(* IEC 61131-3 sources: plcassist-cli/packages/volt-lsp-iec/test-corpus/awa-palletizer/Device/Plc Logic/Application/Library Manager/L_TS2P_TechModulesSynchronizingCamming, 102 files *)

(* ---- L_TS2P_INTERNAL.gvl ---- *)
VAR_GLOBAL
	CDIENUMSTARTVALUE : DINT := 22000;
END_VAR

(* ---- L_TS2M_ITFFLYINGSAWSTATEFMDATA.itf ---- *)
INTERFACE L_TS2M_ITFFLYINGSAWSTATEFMDATA
END_INTERFACE

(* ---- L_TS2M_ITFFLYINGSAWSTATETMDATA.itf ---- *)
INTERFACE L_TS2M_ITFFLYINGSAWSTATETMDATA
END_INTERFACE

METHOD MOVETOPARKPOS : BOOL
VAR_INPUT
	XEXECUTEMOVETOPARKPOS : BOOL;
	LRPARKPOSITION : LREAL := 180;
	EPOSITIONINGDIRECTION : MC_DIRECTION := MC_DIRECTION.mcPositiveDirection;
	LRPOSITIONINGVEL : LREAL := 10;
	LRPOSITIONINGACC : LREAL := 100;
	LRPOSITIONINGDEC : LREAL := 100;
	LRJERK : LREAL := 0;
END_VAR
VAR_OUTPUT
	XBUSY : BOOL;
	XDONE : BOOL;
	XCOMMANDABORTED : BOOL;
END_VAR
VAR_IN_OUT
	AXIS : AXIS_REF;
END_VAR
END_METHOD

(* ---- L_TS2P_ICONNECTORFLEXCAM.itf ---- *)
INTERFACE L_TS2P_ICONNECTORFLEXCAM
END_INTERFACE

(* ---- L_TS2P_ICONNECTORFLYINGSAW.itf ---- *)
INTERFACE L_TS2P_ICONNECTORFLYINGSAW
END_INTERFACE

(* ---- L_TS2P_ICONNECTORSYNCANDCORRECTION.itf ---- *)
INTERFACE L_TS2P_ICONNECTORSYNCANDCORRECTION
END_INTERFACE

(* ---- L_TS2P_ICONNECTORSYNCPOS.itf ---- *)
INTERFACE L_TS2P_ICONNECTORSYNCPOS
END_INTERFACE

(* ---- L_TS2P_IFLEXCAM.itf ---- *)
INTERFACE L_TS2P_IFLEXCAM
END_INTERFACE

METHOD CAM
VAR_INPUT
	ITFTECHMODULE : L_TS2P_IFlexCam;
	XENABLE : BOOL;
	XSYNCCAM : BOOL;
	SCCAMTABLE : MC_CAM_REF;
	LRCYCMASTERPOS : LREAL;
	LRCYCMASTERVEL : LREAL;
	LRCYCMASTERACC : LREAL;
	LRSLAVEPOS : LREAL;
	LRSLAVEVEL : LREAL;
	LRSLAVEACC : LREAL;
	EOFFSETMODEMASTER : L_TS2P_OffsetMode := L_TS2P_OffsetMode.x_zero;
	ESCALINGMODEMASTER : L_TS2P_ScalingMode := L_TS2P_ScalingMode.x_zero;
	EOFFSETMODESLAVE : L_TS2P_OffsetMode := L_TS2P_OffsetMode.x_zero;
	ESCALINGMODESLAVE : L_TS2P_ScalingMode := L_TS2P_ScalingMode.x_zero;
	LRSETOFFSETMASTER : LREAL;
	LRSETOFFSETSLAVE : LREAL;
	LRSETSCALINGMASTER : LREAL;
	LRSETSCALINGSLAVE : LREAL;
	LRPROFGENMASTERVEL : LREAL;
	LRPROFGENMASTERACC : LREAL;
	LRPROFGENMASTERDEC : LREAL;
	LRPROFGENMASTERJERK : LREAL;
	LRPROFGENSLAVEVEL : LREAL;
	LRPROFGENSLAVEACC : LREAL;
	LRPROFGENSLAVEDEC : LREAL;
	LRPROFGENSLAVEJERK : LREAL;
	XPERIODIC : BOOL;
	XCAMCHANGEINSTANT : BOOL;
	XMASTERABSOLUTE : BOOL;
	XSLAVEABSOLUTE : BOOL;
END_VAR
VAR_OUTPUT
	XERROR : BOOL;
	EERRORID : L_IE1P.L_IE1P_Error;
	LRSETPOSOUT : LREAL;
	LRSETVELOUT : LREAL;
	LRSETACCOUT : LREAL;
	LRSETXPOSOUT : LREAL;
	LRSETXVELOUT : LREAL;
	LRSETXACCOUT : LREAL;
	LRSETYPOSOUT : LREAL;
	LRSETYVELOUT : LREAL;
	LRSETYACCOUT : LREAL;
	XENDOFPROFILE : BOOL;
	LRSETOFFSETMASTEROUT : LREAL;
	LRSETOFFSETSLAVEOUT : LREAL;
	LRCONVERTMASTERTOXPOS : LREAL;
	LRCAMPROFILERPOSOUT : LREAL;
	LRCONVERTYTOSLAVEPOS : LREAL;
	XDONE : BOOL;
	XBUSY : BOOL;
END_VAR
END_METHOD

METHOD CAMSEQUENCER
VAR_INPUT
	ITFTECHMODULE : L_TS2P_IFlexCam;
	XENABLE : BOOL;
	XCAMSEQUENCER : BOOL;
	XENDOFPROFILEIN : BOOL;
	CAMTABLE1 : MC_CAM_REF;
	CAMTABLE2 : MC_CAM_REF;
	CAMTABLE3 : MC_CAM_REF;
	CAMTABLE4 : MC_CAM_REF;
	XCAMCHANGEINSTANT : BOOL;
	XLOADCAMTABLE : BOOL;
	WSETCAMTABLE : WORD;
	EMODE : L_TS2P_CamSequenceMode := L_TS2P_CamSequenceMode.CyclicCam1;
END_VAR
VAR_OUTPUT
	XERROR : BOOL;
	EERRORID : L_IE1P_Error;
	CAMTABLEOUT : MC_CAM_REF;
	XCAMTABLEVALID : BOOL;
END_VAR
END_METHOD

METHOD CLUTCH
VAR_INPUT
	ITFTECHMODULE : L_TS2P_IFlexCam;
	XENABLE : BOOL;
	XCLUTCHCLOSE : BOOL;
	ECLUTCHINMODE : L_TS2P_ClutchInMode;
	ECLUTCHOUTMODE : L_TS2P_ClutchOutMode;
	EALLOWEDDIRECTION : L_TB2P_AllowedDirection;
	LRCLUTCHINDIST : LREAL;
	LRCLUTCHOUTDIST : LREAL;
	LRCLUTCHOUTPOSITION : LREAL;
	LRCYCLICMASTERPOS : LREAL;
	LRCYCLICMASTERVEL : LREAL;
	LRCYCLICMASTERACC : LREAL;
	LRCYCLICAXISPOS : LREAL;
	LRCYCLICAXISVEL : LREAL;
	LRCYCLICAXISACC : LREAL;
	ETRAVERSINGRANGE : L_MC1P_TraversingRange;
	LRCYCLELENGTH : LREAL;
END_VAR
VAR_OUTPUT
	XERROR : BOOL;
	EERRORID : L_IE1P.L_IE1P_Error;
	XBUSY : BOOL;
	XDONE : BOOL;
	XSYNCHRONISED : BOOL;
	XACCDECSYNC : BOOL;
	LRSETPOSOUT : LREAL;
	LRSETVELOUT : LREAL;
	LRSETACCOUT : LREAL;
END_VAR
END_METHOD

METHOD HALT : BOOL
VAR_INPUT
	ITFTECHMODULE : L_TS2P_IFlexCam;
	XEXECUTE : BOOL;
	LRDEC : LREAL := 100;
	LRJERK : LREAL := 0;
END_VAR
VAR_OUTPUT
	XBUSY : BOOL;
	XDONE : BOOL;
	XCOMMANDABORTED : BOOL;
END_VAR
VAR_IN_OUT
	AXIS : AXIS_REF;
END_VAR
END_METHOD

METHOD MOVETOPARKPOS : BOOL
VAR_INPUT
	ITFTECHMODULE : L_TS2P_IFlexCam;
	XEXECUTEMOVETOPARKPOS : BOOL;
	EMOVETOPARKPOSMODE : L_TS2P_CamStopMode;
	LRPARKPOSITION : LREAL := 180;
	EPOSITIONINGDIRECTION : L_TS2P_SyncDirection := L_TS2P_SyncDirection.PositiveDirection;
	LRPOSITIONINGVEL : LREAL := 10;
	LRPOSITIONINGACC : LREAL := 100;
	LRPOSITIONINGDEC : LREAL := 100;
	LRJERK : LREAL := 0;
END_VAR
VAR_OUTPUT
	XBUSY : BOOL;
	XDONE : BOOL;
	XCOMMANDABORTED : BOOL;
END_VAR
VAR_IN_OUT
	AXIS : AXIS_REF;
END_VAR
END_METHOD

METHOD POSITIONFOLLOWER
VAR_INPUT
	ITFTECHMODULE : L_TS2P_IFlexCam;
	XENABLE : BOOL;
	LRPOSITION : LREAL;
	LRVELOCITY : LREAL;
	LRACCELERATION : LREAL;
	ESETVALUEMODE : L_MC1P_SetValueMode;
END_VAR
VAR_OUTPUT
	XERROR : BOOL;
	EERRORID : L_IE1P.L_IE1P_Error;
	XBUSY : BOOL;
END_VAR
END_METHOD

METHOD SYNCIN
VAR_INPUT
	ITFTECHMODULE : L_TS2P_IFlexCam;
	XENABLE : BOOL;
	XSYNCIN : BOOL;
	XSYNCPOSRESTORE : BOOL;
	ESYNCMODE : L_TS2P_SyncInMode;
	ESYNCDIRECTION : L_TS2P_SyncDirection;
	LRSYNCVEL : LREAL;
	LRSYNCACC : LREAL;
	LRSYNCDEC : LREAL;
	LRSYNCJERK : LREAL;
	LRPARKPOSITION : LREAL;
	LRCYCLICMASTERPOS : LREAL;
	LRCYCLICMASTERVEL : LREAL;
	LRCYCLICMASTERACC : LREAL;
	LRCYCLICAXISPOS : LREAL;
	LRCYCLICAXISVEL : LREAL;
	LRCYCLICAXISACC : LREAL;
END_VAR
VAR_OUTPUT
	XERROR : BOOL;
	EERRORID : L_IE1P.L_IE1P_Error;
	XBUSY : BOOL;
	XDONE : BOOL;
	XSYNCHRONISED : BOOL;
	XACCDECSYNC : BOOL;
	LRSETPOSOUT : LREAL;
	LRSETVELOUT : LREAL;
	LRSETACCOUT : LREAL;
	LROFFSETSYNCPOS : LREAL;
END_VAR
VAR_IN_OUT
	AXIS : AXIS_REF;
END_VAR
END_METHOD

(* ---- L_TS2P_IFLYINGSAWPROCESSING.itf ---- *)
INTERFACE L_TS2P_IFLYINGSAWPROCESSING
END_INTERFACE

METHOD CLUTCH
VAR_INPUT
	ITFTECHMODULE : L_TS2P_IFlyingSawProcessing;
	XENABLE : BOOL;
	XSYNCVEL : BOOL := FALSE;
	XSYNCPOS : BOOL;
	XSYNCOUTINSTANT : BOOL;
	LRSYNCVEL : LREAL := 10;
	LRSYNCACC : LREAL := 100;
	LRSYNCDEC : LREAL := 100;
	LRSYNCJERK : LREAL := 10000;
	LRCYCMASTERPOS : LREAL;
	LRCYCMASTERVEL : LREAL;
	LRCYCMASTERACC : LREAL;
	LRSETSLAVEPOS : LREAL;
	LRSETSLAVEVEL : LREAL;
	LRSETSLAVEACC : LREAL;
END_VAR
VAR_OUTPUT
	EERRORID : L_IE1P_Error;
	XERROR : BOOL;
	XBUSY : BOOL;
	XDONE : BOOL;
	XACCDECSYNC : BOOL;
	XVELSYNCHRONISED : BOOL;
	XPOSSYNCHRONISED : BOOL;
	LRSETSLAVEPOSOUT : LREAL;
	LRSETSLAVEVELOUT : LREAL;
	LRSETSLAVEACCOUT : LREAL;
	XPROFILERESETTIMEVALID : BOOL;
	LRPROFILERESETTIME : LREAL;
END_VAR
END_METHOD

METHOD EXECUTEGAP
VAR_INPUT
	ITFTECHMODULE : L_TS2P_IFlyingSawProcessing;
	XENABLE : BOOL;
	LRSYNCVEL : LREAL := 10;
	LRSYNCACC : LREAL := 100;
	LRSYNCDEC : LREAL := 100;
	LRSYNCJERK : LREAL := 10000;
	XEXECUTEGAP : BOOL;
	XAUXEXECUTEGAP : BOOL := FALSE;
	LRCYCMASTERPOS : LREAL;
	LRCYCMASTERVEL : LREAL;
	LRCYCMASTERACC : LREAL;
	LRSETSLAVEPOS : LREAL;
	LRSETSLAVEVEL : LREAL;
	LRSETSLAVEACC : LREAL;
END_VAR
VAR_OUTPUT
	EERRORID : L_IE1P_Error;
	XERROR : BOOL;
	XBUSY : BOOL;
	XDONE : BOOL;
	XACCDECSYNC : BOOL;
	XVELSYNCHRONISED : BOOL;
	XPOSSYNCHRONISED : BOOL;
	LRSETSLAVEPOSOUT : LREAL;
	LRSETSLAVEVELOUT : LREAL;
	LRSETSLAVEACCOUT : LREAL;
	XPROFILERESETTIMEVALID : BOOL;
	LRPROFILERESETTIME : LREAL;
END_VAR
END_METHOD

METHOD MARKSTACK_GETMARK
VAR_INPUT
	ITFTECHMODULE : L_TS2P_IFlyingSawProcessing;
	XENABLE : BOOL;
	XGETMARK : BOOL;
	XRESETGETMARK : BOOL;
	XRESETMARKSTACK : BOOL;
	LRCYCSETPOS : LREAL;
	LRCYCSETVEL : LREAL;
END_VAR
VAR_OUTPUT
	XMARKSTACKFULL : BOOL;
	XMARKSTACKEMPTY : BOOL;
	WMARKSINSTACK : WORD;
	XMARKVALID : BOOL;
	LRMARKPOSOUT : LREAL;
END_VAR
END_METHOD

METHOD MARKSTACK_SETMARK
VAR_INPUT
	ITFTECHMODULE : L_TS2P_IFlyingSawProcessing;
	XENABLE : BOOL;
	XSETMARK : BOOL;
	LRMARKPOS : LREAL;
	XRESETMARKSTACK : BOOL;
	LRCYCSETPOS : LREAL;
	LRCYCSETVEL : LREAL;
END_VAR
VAR_OUTPUT
	XMARKSTACKFULL : BOOL;
	XMARKSTACKEMPTY : BOOL;
	WMARKSINSTACK : WORD;
	XNEWMARKRECEIVED : BOOL;
END_VAR
END_METHOD

METHOD POSITIONING
VAR_INPUT
	ITFTECHMODULE : L_TS2P_IFlyingSawProcessing;
	XENABLE : BOOL;
	XMOVETOTARGETPOS : BOOL;
	LRTARGETPOS : LREAL;
	LRPOSITIONINGVEL : LREAL;
	LRPOSITIONINGACC : LREAL;
	LRPOSITIONINGDEC : LREAL;
	LRPOSITIONINGJERK : LREAL;
	LRSETSLAVEPOS : LREAL;
	LRSETSLAVEVEL : LREAL;
	LRSETSLAVEACC : LREAL;
	LRCORRECTTIMEBASE : LREAL := 0;
	LROVERRIDE : LREAL := 1.0;
END_VAR
VAR_OUTPUT
	EERRORID : L_IE1P_Error;
	XERROR : BOOL;
	XBUSY : BOOL;
	XDONE : BOOL;
	XPOSITIONING : BOOL;
	XINPOSITION : BOOL;
	LRSETSLAVEPOSOUT : LREAL;
	LRSETSLAVEVELOUT : LREAL;
	LRSETSLAVEACCOUT : LREAL;
	XPROFILERESETTIMEVALID : BOOL;
	LRPROFILERESETTIME : LREAL;
END_VAR
END_METHOD

(* ---- L_TS2P_ISIGNALFLOW.itf ---- *)
INTERFACE L_TS2P_ISIGNALFLOW
END_INTERFACE

METHOD GET_PSF : POINTER TO L_TS2P_scSF_TM_SyncPosBase
END_METHOD

(* ---- L_TS2P_ISIGNALFLOWFLEXCAM.itf ---- *)
INTERFACE L_TS2P_ISIGNALFLOWFLEXCAM
END_INTERFACE

METHOD GET_PSF : POINTER TO L_TS2P_scSF_TM_SyncPosBase
END_METHOD

(* ---- L_TS2P_ISIGNALFLOWSC.itf ---- *)
INTERFACE L_TS2P_ISIGNALFLOWSC
END_INTERFACE

METHOD GET_PSF : POINTER TO L_TS2P_scSF_TM_SyncAndCorrectionState
END_METHOD

(* ---- L_TS2P_ISTRUCTPROVIDERFLEXCAMHIGH.itf ---- *)
INTERFACE L_TS2P_ISTRUCTPROVIDERFLEXCAMHIGH
END_INTERFACE

METHOD GET_PDATA : POINTER TO L_TS2P_scData_TM_FlexCam
END_METHOD

METHOD GET_PDATASP : POINTER TO L_TS2P_scData_TM_FlexCam
END_METHOD

(* ---- L_TS2P_ISTRUCTPROVIDERFLYINGSAW.itf ---- *)
INTERFACE L_TS2P_ISTRUCTPROVIDERFLYINGSAW
END_INTERFACE

METHOD GET_PDATA : POINTER TO L_TS2M_scData_FlyingSawState
END_METHOD

METHOD GET_PFMDATA : POINTER TO L_TS2M_scData_FM_FlyingSaw
END_METHOD

(* ---- L_TS2P_ISTRUCTPROVIDERSYNCANDCORRECTION.itf ---- *)
INTERFACE L_TS2P_ISTRUCTPROVIDERSYNCANDCORRECTION
END_INTERFACE

METHOD GET_PDATA : POINTER TO L_TS2P_scData_TM_SyncAndCorrectionState
END_METHOD

METHOD GET_PDATASP : POINTER TO L_TS2P_scData_TM_SyncPosBase
END_METHOD

(* ---- L_TS2P_ISTRUCTPROVIDERSYNCPOS.itf ---- *)
INTERFACE L_TS2P_ISTRUCTPROVIDERSYNCPOS
END_INTERFACE

METHOD GET_PDATA : POINTER TO L_TS2P_scData_TM_SyncPosBase
END_METHOD

(* ---- L_TS2P_ISYNCANDCORRECTIONSTATE.itf ---- *)
INTERFACE L_TS2P_ISYNCANDCORRECTIONSTATE
END_INTERFACE

(* ---- L_TS2P_ISYNCPOSBASE.itf ---- *)
INTERFACE L_TS2P_ISYNCPOSBASE
END_INTERFACE

METHOD ADDOFFSET
VAR_INPUT
	ITFTECHMODULE : L_TS2P_ISyncPosBase;
	LRSETPOS : LREAL;
	LRSETVEL : LREAL;
	LRSETOFFSET : LREAL;
	LRSETOFFSETVEL : LREAL;
	ETRAVERSINGRANGE : L_MC1P.L_MC1P_TraversingRange;
	LRCYCLELENGTH : LREAL;
END_VAR
VAR_OUTPUT
	XERROR : BOOL;
	EERRORID : L_IE1P.L_IE1P_Error;
	LRSETPOSOUT : LREAL;
	LRSETVELOUT : LREAL;
END_VAR
END_METHOD

METHOD CLUTCH
VAR_INPUT
	ITFTECHMODULE : L_TS2P_ISyncPosBase;
	XENABLE : BOOL;
	XSYNCIN : BOOL;
	LRSETBASEVELOCITY : LREAL;
	ESYNCMODE : L_TB2P_SyncMode;
	EALLOWEDDIRECTION : L_TB2P_AllowedDirection;
	LRSYNCVEL : LREAL;
	LRSYNCACC : LREAL;
	LRSYNCDEC : LREAL;
	LRSYNCJERK : LREAL;
	LRSYNCINDIST : LREAL;
	LRSYNCOUTDIST : LREAL;
	LRSYNCOUTPOS : LREAL;
	XLOADCLUTCHOFFSET : BOOL;
	LRLOADCLUTCHOFFSET : LREAL;
	LRCYCLICMASTERPOS : LREAL;
	LRCYCLICMASTERVEL : LREAL;
	ETRAVERSINGRANGEMASTER : L_MC1P_TraversingRange;
	LRCYCLELENGTHMASTER : LREAL;
	LRCYCLICAXISPOS : LREAL;
	LRCYCLICAXISVEL : LREAL;
	LRCYCLICAXISACC : LREAL;
	ETRAVERSINGRANGEAXIS : L_MC1P_TraversingRange;
	LRCYCLELENGTHAXIS : LREAL;
END_VAR
VAR_OUTPUT
	XERROR : BOOL;
	EERRORID : L_IE1P.L_IE1P_Error;
	XBUSY : BOOL;
	XDONE : BOOL;
	XSYNCHRONISED : BOOL;
	XACCDECSYNC : BOOL;
	XINBASEVELOCITY : BOOL;
	LRSETPOSOUT : LREAL;
	LRSETVELOUT : LREAL;
	LRSETACCOUT : LREAL;
	LRCLUTCHOFFSETOUT : LREAL;
END_VAR
END_METHOD

METHOD GEARBOX
VAR_INPUT
	ITFTECHMODULE : L_TS2P_ISyncPosBase;
	XENABLE : BOOL;
	LRSETPOSX : LREAL;
	LRSETVELX : LREAL;
	DWNUMERATOR : DWORD;
	DWDENOMINATOR : DWORD;
	LRCYCLELENGTHX : LREAL;
	LRCYCLELENGTHY : LREAL;
	ETRAVERSINGRANGEX : L_MC1P.L_MC1P_TraversingRange;
	ETRAVERSINGRANGEY : L_MC1P.L_MC1P_TraversingRange;
	XLOADGEARBOXPOS : BOOL;
	LRLOADGEARBOXPOS : LREAL;
END_VAR
VAR_OUTPUT
	XERROR : BOOL;
	EERRORID : L_IE1P.L_IE1P_Error;
	LRSETPOSOUT : LREAL;
	LRSETVELOUT : LREAL;
END_VAR
END_METHOD

METHOD OFFSETANDTRIM
VAR_INPUT
	ITFTECHMODULE : L_TS2P_ISyncPosBase;
	XENABLE : BOOL;
	LRSETOFFSET : LREAL;
	XTRIMPOS : BOOL;
	XTRIMNEG : BOOL;
	LRSETTRIMDISTANCE : LREAL;
	ETRIMMODE : L_TS2P_TrimMode;
	XLOADOFFSET : BOOL;
	XRESETTRIMOFFSET : BOOL;
	LRSETVEL : LREAL;
	LRSETACC : LREAL;
	LRSETDEC : LREAL;
	LRSETJERK : LREAL;
	WACTDIRECTION : WORD;
	EALLOWEDDIRECTION : L_TB2P.L_TB2P_AllowedDirection;
	LRCYCMASTERPOS : LREAL;
	LRCYCMASTERVEL : LREAL;
	LRCYCMASTERACC : LREAL;
END_VAR
VAR_OUTPUT
	XERROR : BOOL;
	EERRORID : L_IE1P.L_IE1P_Error;
	XBUSY : BOOL;
	XDONE : BOOL;
	LRSETOFFSETOUTTOTAL : LREAL;
	LRSETOFFSETOUTTOTALVEL : LREAL;
	LRSETOFFSETOUT : LREAL;
	LRSETOFFSETOUTTRIM : LREAL;
END_VAR
END_METHOD

(* ---- GETBOOLEANPROPERTY.fun ---- *)
FUNCTION GETBOOLEANPROPERTY : BOOL
VAR_INPUT
	STKEY : WSTRING;
END_VAR
END_FUNCTION

(* ---- GETCOMPANY.fun ---- *)
FUNCTION GETCOMPANY : WSTRING
END_FUNCTION

(* ---- GETNUMBERPROPERTY.fun ---- *)
FUNCTION GETNUMBERPROPERTY : DINT
VAR_INPUT
	STKEY : WSTRING;
END_VAR
END_FUNCTION

(* ---- GETTEXTPROPERTY.fun ---- *)
FUNCTION GETTEXTPROPERTY : WSTRING
VAR_INPUT
	STKEY : WSTRING;
END_VAR
END_FUNCTION

(* ---- GETTEXTPROPERTY2.fun ---- *)
FUNCTION GETTEXTPROPERTY2 : POINTER TO WSTRING
VAR_INPUT
	STKEY : WSTRING;
END_VAR
END_FUNCTION

(* ---- GETTITLE.fun ---- *)
FUNCTION GETTITLE : WSTRING
END_FUNCTION

(* ---- GETVERSION.fun ---- *)
FUNCTION GETVERSION : VERSION
END_FUNCTION

(* ---- GETVERSIONPROPERTY.fun ---- *)
FUNCTION GETVERSIONPROPERTY : VERSION
VAR_INPUT
	STKEY : WSTRING;
END_VAR
END_FUNCTION

(* ---- L_MB1P_CONVERTPOSTOMODULOPOS.fun ---- *)
FUNCTION L_MB1P_CONVERTPOSTOMODULOPOS : LREAL
VAR_INPUT
	LRPOS : LREAL;
	LRPERIOD : LREAL;
END_VAR
VAR_OUTPUT
	DIREVCOUNTER : DINT;
END_VAR
END_FUNCTION

(* ---- L_MB1P_CONVERTPOSTOMODULOPOSEXTENDED.fun ---- *)
FUNCTION L_MB1P_CONVERTPOSTOMODULOPOSEXTENDED : LREAL
VAR_INPUT
	LRPOS : LREAL;
	LRPERIOD : LREAL;
END_VAR
VAR_OUTPUT
	DIREVCOUNTER : DINT;
END_VAR
END_FUNCTION

(* ---- L_MB1P_CONVERTPOSTOMODULOPOSFMOD.fun ---- *)
FUNCTION L_MB1P_CONVERTPOSTOMODULOPOSFMOD : LREAL
VAR_INPUT
	LRPOS : LREAL;
	LRPERIOD : LREAL;
END_VAR
END_FUNCTION

(* ---- L_MB1P_HLPCALCKOEFPOLY5THORD.fun ---- *)
FUNCTION L_MB1P_HLPCALCKOEFPOLY5THORD : ARRAY [0..5] OF LREAL
VAR_INPUT
	LRYPOSSTART : LREAL;
	LRYVELSTART : LREAL;
	LRYACCSTART : LREAL;
	LRYPOSEND : LREAL;
	LRYVELEND : LREAL;
	LRYACCEND : LREAL;
END_VAR
VAR_OUTPUT
	ALRKOEF : ARRAY [0..5] OF LREAL;
END_VAR
END_FUNCTION

(* ---- L_MB1P_HLPCALCYOFPOLY5THORDBASE.fun ---- *)
FUNCTION L_MB1P_HLPCALCYOFPOLY5THORDBASE : LREAL
VAR_OUTPUT
	LRYPOSSCALED : LREAL;
END_VAR
VAR_IN_OUT
	LRXPOSSCALED : LREAL;
	ALRKOEF : ARRAY [0..5] OF LREAL;
END_VAR
END_FUNCTION

(* ---- L_MB1P_HLPCALCYOFPOLY5THORDSTATE.fun ---- *)
FUNCTION L_MB1P_HLPCALCYOFPOLY5THORDSTATE : LREAL
VAR_INPUT
	LRXPOSSTART : LREAL;
	LRXPOSEND : LREAL := 1;
	LRSETXPOS : LREAL;
	ALRKOEF : ARRAY [0..5] OF LREAL;
END_VAR
VAR_OUTPUT
	LRYPOSSCALED : LREAL;
END_VAR
END_FUNCTION

(* ---- L_MB1P_HLPDELTAVELTIMEEXTENDED.fun ---- *)
FUNCTION L_MB1P_HLPDELTAVELTIMEEXTENDED : BOOL
VAR_INPUT
	LRVELSTART : LREAL;
	LRACCSTART : LREAL;
	LRMAXACC : LREAL;
	LRMAXJERK : LREAL;
END_VAR
VAR_OUTPUT
	LRTIME : LREAL;
	LRDIST : LREAL;
END_VAR
END_FUNCTION

(* ---- L_MB1P_HLPDELTAVELTIMESTATE.fun ---- *)
FUNCTION L_MB1P_HLPDELTAVELTIMESTATE : BOOL
VAR_INPUT
	LRVELSTART : LREAL;
	LRACCSTART : LREAL;
	LRVELTARGET : LREAL;
	LRACCTARGET : LREAL;
	LRMAXACC : LREAL;
	LRMAXDEC : LREAL;
	LRMAXJERK : LREAL;
END_VAR
VAR_OUTPUT
	LRTIME : LREAL;
	LRDIST : LREAL;
END_VAR
END_FUNCTION

(* ---- L_MB1P_HLPDELTAVELTIMETOCONTANTVEL.fun ---- *)
FUNCTION L_MB1P_HLPDELTAVELTIMETOCONTANTVEL : BOOL
VAR_INPUT
	LRACCSTART : LREAL;
	LRMAXJERK : LREAL;
	WMODE : WORD;
END_VAR
VAR_OUTPUT
	LRVEL : LREAL;
	LRTIME : LREAL;
	LRDIST : LREAL;
END_VAR
END_FUNCTION

(* ---- L_MB1P_HLPRESTTIMEFORDISTANCE.fun ---- *)
FUNCTION L_MB1P_HLPRESTTIMEFORDISTANCE : BOOL
VAR_OUTPUT
	LRTIME : LREAL;
END_VAR
VAR_IN_OUT
	LRVELSTART : LREAL;
	LRACCSTART : LREAL;
	LRDIST : LREAL;
END_VAR
END_FUNCTION

(* ---- L_MB1P_MODULOCYCLE.fun ---- *)
FUNCTION L_MB1P_MODULOCYCLE : LREAL
VAR_INPUT
	LRPOSIN : LREAL;
	LRPOSITIONPERIOD : LREAL;
END_VAR
END_FUNCTION

(* ---- L_TS2P_CALCSYNCTIME.fun ---- *)
FUNCTION L_TS2P_CALCSYNCTIME : BOOL
VAR_INPUT
	LRACTMATERIALVEL : LREAL;
	LRACCMAX : LREAL;
	LRJERKSTART : LREAL;
	LRJERKEND : LREAL;
END_VAR
VAR_OUTPUT
	LRACCTIME : LREAL;
	LRACCDIST : LREAL;
END_VAR
END_FUNCTION

(* ---- L_TS2P_CHECK_CAMREFCHANGED.fun ---- *)
FUNCTION L_TS2P_CHECK_CAMREFCHANGED : BOOL
VAR_INPUT
	CAMREFNEW : MC_CAM_REF;
	CAMREFOLD : MC_CAM_REF;
END_VAR
END_FUNCTION

(* ---- L_TS2P_CHECK_CAMREFVALID.fun ---- *)
FUNCTION L_TS2P_CHECK_CAMREFVALID : BOOL
VAR_INPUT
	CAMREF : MC_CAM_REF;
END_VAR
END_FUNCTION

(* ---- _L_MB1P_AXISCONTROLBYPOS.fb ---- *)
FUNCTION_BLOCK _L_MB1P_AXISCONTROLBYPOS
VAR_INPUT
	XENABLE : BOOL;
	LRSETPOSITION : LREAL;
	LRSETVELOCITY : LREAL;
	LRSETACCELERATION : LREAL;
	ESETVALUEMODE : L_MC1P_SetValueMode := L_MC1P_SetValueMode.Pos;
END_VAR
VAR_OUTPUT
	XBUSY : BOOL;
	XCOMMANDABORTED : BOOL;
	XERROR : BOOL;
	EERRORID : L_IE1P_Error;
	LRSETPOSOUT : LREAL;
END_VAR
VAR_IN_OUT
	AXIS : AXIS_REF;
END_VAR
VAR
	LRSETPOSITION_INT : LREAL;
	XENABLE_OLD : BOOL;
	XBUSY_OLD : BOOL;
	ESTATE : L_MB1P_States;
	MC_HALT1 : MC_HALT;
	FB_FOLLOWSETVALUES : L_MC1P_FollowSetValues;
END_VAR
END_FUNCTION_BLOCK

METHOD CALL_ERRORHANDLER
END_METHOD

METHOD CALL_FBMETHODS
END_METHOD

METHOD CALL_FB_FOLLOWSETVALUES
END_METHOD

METHOD CALL_MC_HALT
END_METHOD

METHOD CALL_MC_HALT_INPUT
END_METHOD

METHOD CALL_OUTPUT
END_METHOD

METHOD CALL_RESETCOMMANDS
END_METHOD

METHOD CALL_RESETOUTPUT
END_METHOD

METHOD CALL_STATEMACHINE
END_METHOD

METHOD CALL_S000_CYCLIC
END_METHOD

METHOD CALL_S001_INIT
END_METHOD

METHOD CALL_S002_READY
END_METHOD

METHOD CALL_S999_ERROR
END_METHOD

(* ---- _L_MB1P_AXISCONTROLBYVEL.fb ---- *)
FUNCTION_BLOCK _L_MB1P_AXISCONTROLBYVEL
VAR_INPUT
	XENABLE : BOOL;
	LRSETVELOCITY : LREAL;
END_VAR
VAR_OUTPUT
	XBUSY : BOOL;
	XCOMMANDABORTED : BOOL;
	XERROR : BOOL;
	EERRORID : L_IE1P_Error;
	LRSETVELOUT : LREAL;
END_VAR
VAR_IN_OUT
	AXIS : AXIS_REF;
END_VAR
VAR
	LRSETVELOCITY_INT : LREAL;
	XENABLE_OLD : BOOL;
	XBUSY_OLD : BOOL;
	ESTATE : L_MB1P_States;
	MC_HALT1 : MC_HALT;
	FB_FOLLOWSETVALUES : L_MC1P_FollowSetValues;
END_VAR
END_FUNCTION_BLOCK

METHOD CALL_ERRORHANDLER
END_METHOD

METHOD CALL_FBMETHODS
END_METHOD

METHOD CALL_FB_FOLLOWSETVALUES
END_METHOD

METHOD CALL_MC_HALT
END_METHOD

METHOD CALL_MC_HALT_INPUT
END_METHOD

METHOD CALL_OUTPUT
END_METHOD

METHOD CALL_RESETCOMMANDS
END_METHOD

METHOD CALL_RESETOUTPUT
END_METHOD

METHOD CALL_STATEMACHINE
END_METHOD

METHOD CALL_S000_CYCLIC
END_METHOD

METHOD CALL_S001_INIT
END_METHOD

METHOD CALL_S002_READY
END_METHOD

METHOD CALL_S999_ERROR
END_METHOD

(* ---- GLOBALTEXTLIST.fb ---- *)
FUNCTION_BLOCK GLOBALTEXTLIST
VAR
	M_TEXTLISTFILE : STRING(255);
	_STNAMESPACE : STRING;
END_VAR
END_FUNCTION_BLOCK

(* ---- L_MB1P_CHECKMODULOOVERRUN.fb ---- *)
FUNCTION_BLOCK L_MB1P_CHECKMODULOOVERRUN
VAR_INPUT
	LRSETPOS : LREAL;
	LRSETVEL : LREAL;
	LRPERIOD : LREAL;
END_VAR
VAR_OUTPUT
	XOVERRUNPOS : BOOL;
	XOVERRUNNEG : BOOL;
END_VAR
VAR
	ALRMEM : ARRAY [1..7] OF LREAL;
END_VAR
END_FUNCTION_BLOCK

METHOD CALL_CHECKMODULOOVERRUN
VAR_IN_OUT
	LRSETPOS : LREAL;
	LRSETVEL : LREAL;
	LRPERIOD : LREAL;
	XOVERRUNPOS : BOOL;
	XOVERRUNNEG : BOOL;
	ALRMEM : ARRAY [1..7] OF LREAL;
END_VAR
END_METHOD

(* ---- L_MB1P_CHECKUNLIMITEDOVERRUN.fb ---- *)
FUNCTION_BLOCK L_MB1P_CHECKUNLIMITEDOVERRUN
VAR_INPUT
	LRSETPOS : LREAL;
	LRSETVEL : LREAL;
	LRPERIOD : LREAL;
END_VAR
VAR_OUTPUT
	XOVERRUNPOS : BOOL;
	XOVERRUNNEG : BOOL;
END_VAR
VAR
	ALRMEM : ARRAY [1..7] OF LREAL;
END_VAR
END_FUNCTION_BLOCK

METHOD CALL_CHECKUNLIMITEDOVERRUN
VAR_IN_OUT
	LRSETPOS : LREAL;
	LRSETVEL : LREAL;
	LRPERIOD : LREAL;
	XOVERRUNPOS : BOOL;
	XOVERRUNNEG : BOOL;
	ALRMEM : ARRAY [1..7] OF LREAL;
END_VAR
END_METHOD

(* ---- L_MB1P_CLUTCHEXTENDEDBASE.fb ---- *)
FUNCTION_BLOCK L_MB1P_CLUTCHEXTENDEDBASE EXTENDS L_MC2P_ClutchBasic
VAR_INPUT
	XENABLE : BOOL;
	XCLUTCHCLOSE : BOOL;
	XCLUTCHOPENINSTANT : BOOL;
	ECLUTCHMODE : L_MB1P_ClutchMode := L_MB1P_ClutchMode.ramp_pos;
	ECLUTCHDIRECTION : L_MC2P_ClutchDirection := L_MC2P_ClutchDirection.mcCurrentDirection;
	EDIRECTION : L_MC1P_Direction := 0;
	LRCYCMASTERPOS : LREAL;
	LRCYCMASTERVEL : LREAL;
	LRCYCMASTERACC : LREAL;
	LRCYCSLAVEPOS : LREAL;
	LRCYCSLAVEVEL : LREAL;
	LRCYCSLAVEACC : LREAL;
	LROPENINSTANTDEC : LREAL;
	LRMASTERCLOSEPOS : LREAL;
	LRMASTERCLOSEDIST : LREAL := 100;
	LRSLAVECLOSEDIST : LREAL := 100;
	LRMASTEROPENDIST : LREAL := 100;
	LRSLAVEOPENDIST : LREAL := 100;
	LRSLAVEOPENPOS : LREAL;
	LRCLOSETIME : LREAL := 5;
	LROPENTIME : LREAL := 5;
	LRCLUTCHVEL : LREAL := 100;
	LRCLUTCHACC : LREAL := 1000.0;
	LRCLUTCHDEC : LREAL := 1000.0;
	LRCLUTCHJERK : LREAL := 1000000.0;
	LRVELTOLERANCE : LREAL := 1;
	LRAXESCYCLELENGTH : LREAL := 360;
	EMASTERTRAVERSINGRANGE : L_MC1P_TraversingRange;
	LRCYCLETIME : LREAL := 0.001;
END_VAR
VAR_OUTPUT
	XERROR : BOOL;
	EERRORID : L_IE1P_Error;
	XBUSY : BOOL;
	XDONE : BOOL;
	XSYNCHRONISED : BOOL;
	XCLUTCHACTIVE : BOOL;
	LRSETSLAVEPOSOUT : LREAL;
	LRSETSLAVEVELOUT : LREAL;
	LRSETSLAVEACCOUT : LREAL;
	LRSETSLAVEOFFSETOUT : LREAL;
	LRX0 : LREAL;
	LRX1 : LREAL;
	LRY0 : LREAL;
	LRY1 : LREAL;
	LRX0N : LREAL;
	LRX1N : LREAL;
	LRY0N : LREAL;
	LRY1N : LREAL;
	LRX0P : LREAL;
	LRX1P : LREAL;
	LRY0P : LREAL;
	LRY1P : LREAL;
END_VAR
VAR
	EAXESTRAVERSINGRANGE_INT : L_MC1P_TraversingRange;
	ECLUTCHMODE_INT : L_MB1P_ClutchMode;
	ECLUTCHDIRECTION_INT : L_MB1P_ClutchDirection;
	LRSETSLAVEOFFSET_CLUTCHREL : LREAL;
	LRSETSLAVEOFFSET_INT : LREAL;
	LRSETMASTEROFFSET_OVERRUN : LREAL;
	LRCYCLETIME_INT : LREAL;
	XCLUTCHOPENINSTANT_ACTIVE : BOOL;
	LROPENINSTANTDEC_INT : LREAL;
	XCLUTCHBASICENABLE : BOOL;
	LRTEMP : LREAL;
	LRDELTASETENDPOS : LREAL;
	LRDELTASETENDPOS_OLD : LREAL;
	LRDELTASETENDPOS_OLD2 : LREAL;
	XCLUTCHMASTERVELPOSITIVE : BOOL;
	XMASTERREVERSING : BOOL;
	XCLUTCHBASIC_EXECUTE_OLD : BOOL;
	XCLUTCHCLOSE_OLD : BOOL;
	XCLUTCHOPENINSTANT_OLD : BOOL;
	XBUSY_OLD : BOOL;
	XENABLE_OLD : BOOL;
	LRCYCMASTERPOS_OLD : LREAL;
	LRMASTERVELADD : LREAL;
	LRMASTERVELADDSYNC : LREAL;
	LRSLAVESTARTPOS : LREAL;
	LRMASTERCLOSEPOS_INT : LREAL;
	LRMASTERCLOSEDIST_INT : LREAL;
	LRSLAVECLOSEDIST_INT : LREAL;
	LRSLAVEOPENDIST_INT : LREAL;
	LRSLAVEOPENPOS_INT : LREAL;
	XSYNCMODEIN_INT : BOOL;
	LRCLUTCHTIME : LREAL;
	XCLUTCHPOSMODE_INT : BOOL := TRUE;
	LRCLUTCHVEL_INT : LREAL := 100;
	LRCLUTCHACC_INT : LREAL := 1000.0;
	LRCLUTCHDEC_INT : LREAL := 1000.0;
	LRCLUTCHJERK_INT : LREAL := 1000000.0;
	EMASTERDIRECTION_INT : L_MC2P_ClutchDirection;
	IMASTERMOVEMENTTYPE_INT : INT;
	XREVERSEALLOWED_INT : BOOL;
	XPERIODIC_INT : BOOL;
	LRSLAVEJERK : LREAL;
	ESTATE : L_MB1P_States := L_MB1P_States.INIT;
	XSTATEENTRY : BOOL;
	XSETPARAGAIN : BOOL;
	XERROR_LOCK : BOOL;
	EERRORID_LOCK : L_IE1P_Error;
	LRTOLERANCE : LREAL;
	ICYCLECNTAFTEREXECUTE : INT;
	XRESTART_INT : BOOL;
	SCCYCMASTER : L_MC2P_AxisProfile;
	SCCYCSLAVE : L_MC2P_AxisProfile;
	SCSETSLAVEOUT : L_MC2P_AxisProfile;
	SCSETSLAVEOUT_OLD : L_MC2P_AxisProfile;
	PSCSETSLAVEOUT : POINTER TO L_MC2P_AxisProfile;
	EMASTERDIRECTION : L_MC2P_ClutchDirection;
	XCLUTCHBASIC_DONE : BOOL;
	XCLUTCHBASIC_WARNINGCANTPREVENTREVERSE : BOOL;
	XCLUTCHBASIC_ERROR : BOOL;
	ECLUTCHBASIC_ERRORIDCLUTCH : L_IE1P_Error;
	XCLUTCHBASIC_BUSY : BOOL;
	XCLUTCHBASIC_CLUTCHACTIVE : BOOL;
	XCLUTCHBASIC_PERIODIC : BOOL;
	XCLUTCHBASIC_REVERSEALLOWED : BOOL;
	ECLUTCHBASIC_MASTERAXISTYPE : L_MC1P_TraversingRange;
	XCLUTCHBASIC_EXECUTE : BOOL;
	FB_CHECKMODULOOVERRUN : L_MB1P_CheckModuloOverrun;
	XHALT_OLD : BOOL;
	XHALTBUSYINT : BOOL;
	XHALTDONEINT : BOOL;
	XSIMPLEFUNRAMPSLAVEDIST : BOOL := TRUE;
	LRSETSLAVEOFFSET_CLUTCHRELENTRY : LREAL;
	XRAMPDISTABSVIALINEAR : BOOL;
	XCLUTCHBASIC_BUSY_OLD : BOOL;
	XCLUTCHMASTERVELPOSITIVE_OLD : BOOL;
	XMASTERINSIDEXSIZE : BOOL;
	XMASTERINSIDEXSIZE_OLD : BOOL;
	XMASTERINSIDEXSIZEP : BOOL;
	XMASTERINSIDEXSIZEP_OLD : BOOL;
	XMASTERINSIDEXSIZEN : BOOL;
	XMASTERINSIDEXSIZEN_OLD : BOOL;
	XCLUTCHDIRECTIONPOSITIVE : BOOL;
	ALRKOEF : ARRAY [0..5] OF LREAL;
	LRXFACTORN : LREAL;
	LRYFACTORN : LREAL;
	LRSETSLAVEOFFSET_CLUTCHRELN : LREAL;
	LRXFACTORP : LREAL;
	LRYFACTORP : LREAL;
	LRSETSLAVEOFFSET_CLUTCHRELP : LREAL;
	LRXFACTOR : LREAL;
	LRYFACTOR : LREAL;
	LRXSCALED : LREAL;
	LRYSCALED : LREAL;
	LRYSCALED_OLD : LREAL;
	LRYSCALEDDIFF : LREAL;
	LRSETYPOS : LREAL;
	LRSETYPOS_OLD : LREAL;
	LRSETYVEL : LREAL;
	LRSETYVEL_OLD : LREAL;
	LRSETYACC : LREAL;
	XCLUTCHDIRECTIONPOSITIVE_OLD : BOOL;
	LRMASTERCYCLELENGTH : LREAL;
	LRDUMMY : LREAL;
	LRCYCMASTERVEL_OLD : LREAL;
	WRAMPVELLACCSTEPPER : WORD;
	XNOREVERSEACTIVE : BOOL;
	XHALT_BUSY : BOOL;
	XHALT_DONE : BOOL;
	XSLAVEHALT : BOOL;
	C_ALRKOEF_SYNCIN : ARRAY [0..5] OF LREAL := [0, 0, 0, 1, -0.5, 0];
	C_ALRKOEF_SYNCOUT : ARRAY [0..5] OF LREAL := [0, 1, 0, -1, 0.5, 0];
END_VAR
END_FUNCTION_BLOCK

METHOD CALL_ALLOCPOINTADR
END_METHOD

METHOD CALL_CLUTCHCLOSEMODE
END_METHOD

METHOD CALL_CLUTCHOPENMODE
END_METHOD

METHOD CALL_ERRORHANDLER
END_METHOD

METHOD CALL_FBMETHODS
END_METHOD

METHOD CALL_FB_CHECKMODULOOVERRUN
END_METHOD

METHOD CALL_FB_CLUTCHBASIC
END_METHOD

METHOD CALL_FB_CLUTCHBASIC_INPUTSMASTER
END_METHOD

METHOD CALL_FB_CLUTCHBASIC_OPENINSTANT
END_METHOD

METHOD CALL_FB_CLUTCHBASIC_RAMPABS
END_METHOD

METHOD CALL_FB_CLUTCHBASIC_RAMPABS_TARGETPOS
END_METHOD

METHOD CALL_FB_CLUTCHBASIC_RAMPPOS
END_METHOD

METHOD CALL_FB_CLUTCHBASIC_RAMPREL
END_METHOD

METHOD CALL_FB_CLUTCHBASIC_RAMPSLAVEDIST
END_METHOD

METHOD CALL_FB_CLUTCHBASIC_RAMPTIME
END_METHOD

METHOD CALL_FB_CLUTCHBASIC_RAMPVELLACC
END_METHOD

METHOD CALL_FB_CLUTCHBASIC_RELATIVE
END_METHOD

METHOD CALL_MODULOTOLINEARMASTERPOS
END_METHOD

METHOD CALL_OUTPUT
END_METHOD

METHOD CALL_RAMPRELDIESTREL_CALCCOEFX0X1Y0Y1
END_METHOD

METHOD CALL_RAMPRELDISTABS_CALCCOEFX0X1Y0Y1
END_METHOD

METHOD CALL_RAMPRELDISTABS_CORRX0X1FORMODULOMASTER
END_METHOD

METHOD CALL_RAMPSLAVEDIST_ABS
END_METHOD

METHOD CALL_RAMPSLAVEDIST_REL
END_METHOD

METHOD CALL_RAMPSLAVEDIST_SETYPOSOUT
END_METHOD

METHOD CALL_RESETCLUTCH
END_METHOD

METHOD CALL_RESETCOMMANDS
END_METHOD

METHOD CALL_RESETOUTPUT
END_METHOD

METHOD CALL_SETCLUTCHCLOSEPAR
END_METHOD

METHOD CALL_SETCLUTCHCLOSEPAR_OLD
END_METHOD

METHOD CALL_SETCLUTCHOPENPAR
END_METHOD

METHOD CALL_SETCLUTCHOPENPAR_OLD
END_METHOD

METHOD CALL_STATEMASHINE
END_METHOD

METHOD SET_CLUTCHOFFSET : BOOL
VAR_INPUT
	LRIN : LREAL := 0;
END_VAR
END_METHOD

METHOD SLAVEHALT
VAR_INPUT
	XHALT : BOOL;
	SCACTSLAVE : L_MC2P_AxisProfile;
	LRMAXVELDIFF : LREAL;
	LRMAXACC : LREAL;
	LRMAXDEC : LREAL;
	LRJERK : LREAL;
	LRCYCLETIME : LREAL;
END_VAR
VAR_OUTPUT
	SCOUTPUTSLAVE : L_MC2P_AxisProfile;
	XBUSY : BOOL;
	XDONE : BOOL;
	XERROR : BOOL;
	EERRORID : L_IE1P_Error;
END_VAR
END_METHOD

METHOD CALL_S000_CYCLIC
END_METHOD

METHOD CALL_S001_INIT
END_METHOD

METHOD CALL_S010_READY
END_METHOD

METHOD CALL_S100_CLUTCH_CLOSE
END_METHOD

METHOD CALL_S200_SYNCHRON
END_METHOD

METHOD CALL_S300_CLUTCH_OPEN
END_METHOD

METHOD CALL_S998_ERROR
END_METHOD

(* ---- L_MB1P_GEARBOXPOSITION.fb ---- *)
FUNCTION_BLOCK L_MB1P_GEARBOXPOSITION EXTENDS L_MB1P_GearboxPositionBase
VAR_IN_OUT
	AXISX : AXIS_REF;
	AXISY : AXIS_REF;
END_VAR
END_FUNCTION_BLOCK

METHOD CALL_ERRORHANDLER
END_METHOD

(* ---- L_MB1P_GEARBOXPOSITIONBASE.fb ---- *)
FUNCTION_BLOCK L_MB1P_GEARBOXPOSITIONBASE
VAR_INPUT
	XENABLE : BOOL;
	LRPOSX : LREAL;
	DWNUMERATOR : DWORD := 1;
	DWDENOMINATOR : DWORD := 1;
	XLOADPOSY : BOOL;
	LRLOADPOSY : LREAL;
	LNLOADPOSYRESIDUAL : LINT;
END_VAR
VAR_OUTPUT
	LRPOSY : LREAL;
	LRVELY : LREAL;
	LNACTPOSYRESIDUAL : LINT;
	XERROR : BOOL := FALSE;
	EERRORID : L_IE1P_Error := 0;
END_VAR
VAR
	XENABLE_OLD : BOOL := FALSE;
	XINITDONE : BOOL := FALSE;
	LNPOSX : LINT := 0;
	LNPOSY : LINT := 0;
	LNPOSXOLD : LINT := 0;
	LNPOSXDIFF : LINT := 0;
	LNPOSYDIFF : LINT := 0;
	LNPOSYOLD : LINT := 0;
	LNRES_GEARBOX : LINT := 0;
	LRLENX : LREAL;
	LRLENY : LREAL;
	LRLENXOLD : LREAL;
	LRLENYOLD : LREAL;
	LRTASKCYCLE : LREAL;
	LRPOSYOLD : LREAL;
	LRGEARFACTOR : LREAL;
	DWGEARFACTOR : DWORD;
	LIAUFLOESUNG : LINT;
END_VAR
END_FUNCTION_BLOCK

METHOD CALL_S000_CYCLIC
END_METHOD

METHOD CALL_ERRORHANDLER
END_METHOD

METHOD CALL_RESET
END_METHOD

METHOD L_HLPMODULOADD : LREAL
VAR_INPUT
	LRINPUT : LINT;
	LROFFSET : LINT;
	LRLENGHT : LINT;
END_VAR
END_METHOD

METHOD L_HLPMODULODIFF : LREAL
VAR_INPUT
	LRDIFF : LINT;
	LRLEN : LINT;
END_VAR
END_METHOD

METHOD L_HLPMULDIV : LREAL
VAR_INPUT
	LNINPUT : LINT;
	DWNUMERATOR : DWORD;
	DWDENOMINATOR : DWORD;
	PLNRES : POINTER TO LINT;
END_VAR
END_METHOD

(* ---- L_MB1P_GEARBOXPOSITIONINPUT.fb ---- *)
FUNCTION_BLOCK L_MB1P_GEARBOXPOSITIONINPUT EXTENDS L_MB1P_GearboxPositionBase
VAR_INPUT
	LRCYCLELENGTHX : LREAL;
	LRCYCLELENGTHY : LREAL;
END_VAR
END_FUNCTION_BLOCK

(* ---- L_MB1P_POSPROFILERCLUTCH.fb ---- *)
FUNCTION_BLOCK L_MB1P_POSPROFILERCLUTCH
VAR_INPUT
	XENABLE : BOOL;
	XSYNCPOS : BOOL;
	XEXECUTEGAP : BOOL;
	XAUXEXECUTEGAP : BOOL;
	LRTASKCYCLETIME : LREAL := 0.001;
	LRSLAVESYNCOUTPOS : LREAL;
	LRCYCMASTERPOS : LREAL;
	LRCYCMASTERVEL : LREAL;
	LRCYCMASTERACC : LREAL;
	LRSETSLAVEPOS : LREAL;
	LRSETSLAVEVEL : LREAL;
	LRSETSLAVEACC : LREAL;
	LRJERK : LREAL := 10000;
	LRMAXACC : LREAL := 100;
	LRMAXDEC : LREAL := 100;
	LRMAXVEL : LREAL := 10;
END_VAR
VAR_OUTPUT
	XBUSY : BOOL;
	XDONE : BOOL;
	XACCDECSYNC : BOOL;
	XPOSSYNCHRONISED : BOOL;
	XERROR : BOOL;
	EERRORID : WORD;
	LRSETSLAVEPOSOUT : LREAL;
	LRSETSLAVEVELOUT : LREAL;
	LRSETSLAVEACCOUT : LREAL;
	XPROFILERESETTIMEVALID : BOOL;
	LRPROFILERESETTIME : LREAL;
END_VAR
VAR
	FB_POSPROFILERPOS : L_MC1P_PosProfiler;
	SCPROFILEPARAMETER : L_MC1P_ProfileParameter;
	WSTEPPER : WORD;
	XEXECUTEPOSPROFILER : BOOL;
	LRSLAVESYNCOUTPOS_INT : LREAL;
	XAUXEXECUTEPROFILE : BOOL;
	XEXECUTEPROFILE : BOOL;
	LRSETPOSPROFILER : LREAL;
	LRSETACCPROFILER : LREAL;
	LRSETVELPROFILER : LREAL;
	LRCYCMASTERPOS_INT : LREAL;
	LRCYCMASTERVEL_INT : LREAL;
	LRCYCMASTERACC_INT : LREAL;
	XPOSSYNCHRONISED_INT : BOOL;
	XEXECUTEGAPOLD : BOOL;
	XAUXEXECUTEGAPOLD : BOOL;
	XENABLEOLD : BOOL;
	LRCYCMASTERPOS_OLD : LREAL;
	LRTOLERANCE : LREAL;
END_VAR
END_FUNCTION_BLOCK

METHOD CALL_ERRORHANDLER
END_METHOD

METHOD CALL_FBMETHODES
END_METHOD

METHOD CALL_FB_POSPROFILERPOS
END_METHOD

METHOD CALL_FB_POSPROFILERPOSINPUTS
END_METHOD

METHOD CALL_OUTPUTS
END_METHOD

METHOD CALL_PROFILEPARAMETER
END_METHOD

METHOD CALL_RESETCOMMANDS
END_METHOD

METHOD CALL_RESETOUTPUTS
END_METHOD

METHOD CALL_STATEMACHINE
END_METHOD

(* ---- L_MB1P_POSPROFILERCLUTCHHIGH.fb ---- *)
FUNCTION_BLOCK L_MB1P_POSPROFILERCLUTCHHIGH EXTENDS L_MB1P_PosProfilerClutchState
VAR_INPUT
	XSYNCVEL : BOOL;
END_VAR
VAR_OUTPUT
	XVELSYNCHRONISED : BOOL;
END_VAR
VAR
	WSTEPPER_OLD : WORD;
	XSYNCVEL_OLD : BOOL;
	LRCYCMASTERPOSOUT : LREAL;
	LRCYCMASTERVELOUT : LREAL;
	LRCYCMASTERACCOUT : LREAL;
	LRMASTEROFFSET_INT : LREAL;
	LRSETSLAVEACCOUT_OLD : LREAL;
	LRSETSLAVEPOSOUT_OLD : LREAL;
	LRSETSLAVEPOSOUT_2OLD : LREAL;
END_VAR
END_FUNCTION_BLOCK

METHOD CALL_CALCTARGETPOS
VAR_INPUT
	LRTARGETPOS : LREAL;
END_VAR
END_METHOD

METHOD CALL_CALCLRCYCMASTERPOS
END_METHOD

METHOD CALL_OUTPUTS
END_METHOD

METHOD CALL_PROFILEPARAMETER
END_METHOD

METHOD CALL_STATEMACHINE
END_METHOD

(* ---- L_MB1P_POSPROFILERCLUTCHSTATE.fb ---- *)
FUNCTION_BLOCK L_MB1P_POSPROFILERCLUTCHSTATE EXTENDS L_MB1P_PosProfilerClutch
VAR_INPUT
	XSYNCOUTINSTANT : BOOL;
	XMOVETOTARGETPOS : BOOL;
	LRCORRECTTIMEBASE : LREAL := 0;
	LRTARGETPOS : LREAL;
	EDIRECTION : L_MC2P_ClutchDirection := L_MC2P_ClutchDirection.mcCurrentDirection;
	LRAXESCYCLELENGTH : LREAL := 360;
	EAXESTRAVERSINGRANGE : L_MC1P_TraversingRange;
	LRPOSITIONINGJERK : LREAL;
	LRPOSITIONINGACC : LREAL;
	LRPOSITIONINGDEC : LREAL;
	LRPOSITIONINGVEL : LREAL;
	LRSYNCOUTINSTANTJERK : LREAL;
	LRSYNCOUTINSTANTDEC : LREAL;
	ROVERRIDEVEL : REAL := 1.0;
	ROVERRIDEACC : REAL := 1.0;
	ROVERRIDEDEC : REAL := 1.0;
END_VAR
VAR_OUTPUT
	XREVERSING : BOOL;
	XPOSITIONING : BOOL;
	XINPOSITION : BOOL;
END_VAR
VAR
	XREVERSING_INT : BOOL;
	LRCORRECTTIMEBASE_INT : LREAL := 0;
	WMODE : WORD;
	XSYNCOUTINSTANT_OLD : BOOL;
	XMOVETOTARGETPOS_OLD : BOOL;
	XPOSMODE_INT : BOOL;
	LRTASKCYCLETIME_INT : LREAL;
	LRAXESCYCLELENGTH_INT : LREAL;
	LRTARGETPOS_INT : LREAL;
	LRTARGETPOS_LOCK : LREAL;
	LRTOLERANCEVEL : LREAL;
	LRTOLERANCEACC : LREAL;
	LRACCDIST : LREAL;
	XVELTRACE : BOOL;
	WVELTRACESTEPPER : WORD;
	LRSETACC_PROFILERPOS : LREAL;
	LRPOSPROFILERSPEED_ABS : LREAL;
	WREVERSINGVELMODE : WORD;
	LRVELZERROTOLERANZ : LREAL;
	LRSETSLAVEVELOUT_OLD : LREAL;
END_VAR
END_FUNCTION_BLOCK

METHOD CALL_CALCTARGETPOS
VAR_INPUT
	LRTARGETPOS : LREAL;
END_VAR
END_METHOD

METHOD CALL_CALCTOLERANCE
END_METHOD

METHOD CALL_CALCLRCYCMASTERPOS
END_METHOD

METHOD CALL_ERRORHANDLER
END_METHOD

METHOD CALL_FBMETHODES
END_METHOD

METHOD CALL_FB_POSPROFILERPOS
END_METHOD

METHOD CALL_FB_POSPROFILERPOSINPUTS
END_METHOD

METHOD CALL_OUTPUTS
END_METHOD

METHOD CALL_PROFILEPARAMETER
END_METHOD

METHOD CALL_PROFILEPARAMETERACCDECINMODE2
END_METHOD

METHOD CALL_RESETCOMMANDS
END_METHOD

METHOD CALL_RESETOUTPUTS
END_METHOD

METHOD CALL_STATEMACHINE
END_METHOD

(* ---- L_MB1P_STACK.fb ---- *)
FUNCTION_BLOCK L_MB1P_STACK
VAR_INPUT
	XENABLE : BOOL;
	XLOADTPPOS : BOOL;
	XLOADCYCSETPOS : BOOL;
	XTAKEPOS : BOOL;
	LRTPPOS : LREAL;
	LRCYCSETPOS : LREAL;
	LRCYCSETVEL : LREAL;
	LRPERIOD : LREAL;
	LRMINTPDIST : LREAL;
END_VAR
VAR_OUTPUT
	XBUSY : BOOL;
	XSTACKISFULL : BOOL;
	XSTACKISEMPTY : BOOL;
	LRPOSOUT : LREAL;
	LRDISTOUT : LREAL;
	LRSETDISTOUT : LREAL;
	XPOSPERIODOVERRUNPOS : BOOL;
	XPOSPERIODOVERRUNNEG : BOOL;
	UISTACKSTARTPOS : UINT := 0;
	UISTACKFILLSTATE : UINT := 0;
	ALRSTACKSAVEPOS : ARRAY [1..gc_uiStackLength] OF LREAL;
	AUIPERIODCNTRPOS : ARRAY [1..gc_uiStackLength] OF UINT;
	UIPERIODCNTR : UINT;
	LRTPDIST : LREAL;
	XPOSRECEIVED : BOOL;
	XPOSOUTOFWINDOW : BOOL;
	XWINDOWOPEN : BOOL;
END_VAR
VAR
	XSTACKVALUEVALID : BOOL;
	LRLATESTSAVEPOS : LREAL;
	UILATESTPERIODCNTRPOS : UINT;
	UICTR : UINT := 0;
	UIVARTEMP : UINT;
	XENABLE_OLD : BOOL;
	XLOADTPPOS_OLD : BOOL;
	XLOADCYCSETPOS_OLD : BOOL;
	XTAKEPOS_OLD : BOOL;
	XFIRSTLOADPOS : BOOL;
	LRCYCSETPOS_SAVE : LREAL;
	LRSETPOSDIFF : LREAL;
	XTAKEPOS_ACTIVE : BOOL;
	LRTEMPDIST : LREAL;
	LRCYCSETPOS_OLD : LREAL;
	FB_CHECKMODULOOVERRUN : L_MB1P_CheckModuloOverrun;
	GC_UISTACKLENGTH : UINT := 100;
END_VAR
END_FUNCTION_BLOCK

METHOD CALL_CNTRMODULOOVERRUN
VAR_IN_OUT
	LRCYCSETPOS : LREAL;
END_VAR
END_METHOD

METHOD CALL_FB_CHECKMODULOOVERRUN
VAR_IN_OUT
	LRCYCSETPOS : LREAL;
	LRCYCSETVEL : LREAL;
END_VAR
END_METHOD

METHOD CALL_RESETCOMMANDS
END_METHOD

METHOD CALL_RESETOUTPUT
END_METHOD

METHOD CALL_STACK
END_METHOD

METHOD CALL_STACK_LOADPOS
VAR_IN_OUT
	LRCYCPOS : LREAL;
	LRLOADPOS : LREAL;
END_VAR
END_METHOD

METHOD CALL_STACK_TAKEPOS
VAR_IN_OUT
	LRCYCPOS : LREAL;
END_VAR
END_METHOD

METHOD FUN_PERIODCNTRDIFF : LREAL
VAR_INPUT
	UIDIFF : UINT;
END_VAR
VAR_OUTPUT
	IOUT : INT;
END_VAR
END_METHOD

METHOD GET_LRLATESTDIST : LREAL
VAR_IN_OUT
	LRCYCPOS : LREAL;
END_VAR
END_METHOD

METHOD GET_LRTAKEPOS : LREAL
VAR_IN_OUT
	LRCYCPOS : LREAL;
END_VAR
END_METHOD

METHOD REVOKETAKEPOS
END_METHOD

METHOD SET_CYCSETPOS
VAR_IN_OUT
	LRCYCPOS : LREAL;
END_VAR
END_METHOD

METHOD SET_TPPOS
VAR_IN_OUT
	LRCYCPOS : LREAL;
	LRLOADTPPOS : LREAL;
END_VAR
END_METHOD

(* ---- L_MB1P_STACK_FLYINGSAW.fb ---- *)
FUNCTION_BLOCK L_MB1P_STACK_FLYINGSAW
VAR_INPUT
	XENABLE : BOOL;
	XLOADTPPOS : BOOL;
	XLOADCYCSETPOS : BOOL;
	XTAKEPOS : BOOL;
	LRTPPOS : LREAL;
	LRCYCSETPOS : LREAL;
	LRCYCSETVEL : LREAL;
	LRPERIOD : LREAL;
	LRMINTPDIST : LREAL;
END_VAR
VAR_OUTPUT
	XBUSY : BOOL;
	XSTACKISFULL : BOOL;
	XSTACKISEMPTY : BOOL;
	LRPOSOUT : LREAL;
	LRDISTOUT : LREAL;
	LRSETDISTOUT : LREAL;
	XPOSPERIODOVERRUNPOS : BOOL;
	XPOSPERIODOVERRUNNEG : BOOL;
	UISTACKSTARTPOS : UINT := 0;
	UISTACKFILLSTATE : UINT := 0;
	ALRSTACKSAVEPOS : ARRAY [1..gc_uiStackLength] OF LREAL;
	AUIPERIODCNTRPOS : ARRAY [1..gc_uiStackLength] OF UINT;
	UIPERIODCNTR : UINT;
	LRTPDIST : LREAL;
	XPOSRECEIVED : BOOL;
	XPOSOUTOFWINDOW : BOOL;
	XWINDOWOPEN : BOOL;
END_VAR
VAR
	XSTACKVALUEVALID : BOOL;
	LRLATESTSAVEPOS : LREAL;
	UILATESTPERIODCNTRPOS : UINT;
	UICTR : UINT := 0;
	UIVARTEMP : UINT;
	XENABLE_OLD : BOOL;
	XLOADTPPOS_OLD : BOOL;
	XLOADCYCSETPOS_OLD : BOOL;
	XTAKEPOS_OLD : BOOL;
	XFIRSTLOADPOS : BOOL;
	LRCYCSETPOS_SAVE : LREAL;
	LRSETPOSDIFF : LREAL;
	XTAKEPOS_ACTIVE : BOOL;
	LRTEMPDIST : LREAL;
	LRCYCSETPOS_OLD : LREAL;
	FB_CHECKMODULOOVERRUN : L_MB1P_CheckUnlimitedOverrun;
	GC_UISTACKLENGTH : UINT := 100;
END_VAR
END_FUNCTION_BLOCK

METHOD CALL_CNTRMODULOOVERRUN
VAR_IN_OUT
	LRCYCSETPOS : LREAL;
END_VAR
END_METHOD

METHOD CALL_FB_CHECKMODULOOVERRUN
VAR_IN_OUT
	LRCYCSETPOS : LREAL;
	LRCYCSETVEL : LREAL;
END_VAR
END_METHOD

METHOD CALL_RESETCOMMANDS
END_METHOD

METHOD CALL_RESETOUTPUT
END_METHOD

METHOD CALL_STACK
END_METHOD

METHOD CALL_STACK_LOADPOS
VAR_IN_OUT
	LRCYCPOS : LREAL;
	LRLOADPOS : LREAL;
END_VAR
END_METHOD

METHOD CALL_STACK_TAKEPOS
VAR_IN_OUT
	LRCYCPOS : LREAL;
END_VAR
END_METHOD

METHOD FUN_PERIODCNTRDIFF : LREAL
VAR_INPUT
	UIDIFF : UINT;
END_VAR
VAR_OUTPUT
	IOUT : INT;
END_VAR
END_METHOD

METHOD GET_LRLATESTDIST : LREAL
VAR_IN_OUT
	LRCYCPOS : LREAL;
END_VAR
END_METHOD

METHOD GET_LRTAKEPOS : LREAL
VAR_IN_OUT
	LRCYCPOS : LREAL;
END_VAR
END_METHOD

METHOD REVOKETAKEPOS
END_METHOD

METHOD SET_CYCSETPOS
VAR_IN_OUT
	LRCYCPOS : LREAL;
END_VAR
END_METHOD

METHOD SET_TPPOS
VAR_IN_OUT
	LRCYCPOS : LREAL;
	LRLOADTPPOS : LREAL;
END_VAR
END_METHOD

(* ---- L_MC2A_FINDCAMXVALUE.fb ---- *)
FUNCTION_BLOCK L_MC2A_FINDCAMXVALUE
VAR_INPUT
	LRCAMYPOSIN : LREAL;
	LRACTYPOSIN : LREAL;
	LRCYCLELENGTHX : LREAL := 360.0;
	LRCYCLELENGTHY : LREAL := 360.0;
END_VAR
VAR_OUTPUT
	LRCAMXPOSOUT : LREAL;
	LRYDIFFERENCE : LREAL;
	XBUSY : BOOL;
	XDONE : BOOL;
	XERROR : BOOL;
	EERRORID : L_IE1P_ERROR;
END_VAR
END_FUNCTION_BLOCK

METHOD METH_ADDOFFSETCYCLIC : LREAL
VAR_INPUT
	LRSETPOS : LREAL;
	LRSETOFFSET : LREAL;
	LRCYCLELENGTH : LREAL;
END_VAR
END_METHOD

METHOD METH_SHORTESTWAY : LREAL
VAR_INPUT
	LRSETPOS : LREAL;
	LRACTPOS : LREAL;
	LRCYCLELENGTH : LREAL;
END_VAR
END_METHOD

(* ---- L_TS2M_FM_FLYINGSAWSTATE.fb ---- *)
FUNCTION_BLOCK L_TS2M_FM_FLYINGSAWSTATE EXTENDS L_TB2M_FM_Base
VAR_INPUT
	ETMSTATE_EXT : L_TB2P_States;
	AXIS : REFERENCE TO AXIS_REF;
	ITFSTRUCTPROVIDER : L_TS2P_IStructProviderFlyingSaw;
	MASTERVALUES : L_MC1P_IAXIS_REF_MASTERVALUES;
	XSTARTFLYINGSAW : BOOL;
	XSYNCININSTANT : BOOL;
	XEXECUTENEXTCUT : BOOL;
	XEXECUTEGAP : BOOL;
	XSETCUTTINGLENGTHINSTANT : BOOL;
	LRCUTTINGLENGTH : LREAL;
	LRSYNCOVERRIDE : LREAL := 1;
	XSETMATERIALCOUNTER : BOOL;
	XRESUMETARGETPOS : BOOL;
	XRESETMARKSTACK : BOOL;
	PSCTPRECDATA_MARKSENSOR : POINTER TO L_MC1P.L_MC1P_TpReceiveData;
END_VAR
VAR_OUTPUT
	EFM_STATE : L_TB2P_States;
	XSYNCHRONISED : BOOL;
	XACCDECSYNC : BOOL;
	XINPOSITION : BOOL;
	XPOSITIONING : BOOL;
	LRMATERIALCOUNTER : LREAL;
	LRTARGETPOS : LREAL;
	LRCUTGAP : LREAL;
	LRACTIVECUTTINGLENGTH : LREAL;
	WMARKSINSTACK : WORD;
END_VAR
VAR
	ITFFMDATA : L_TS2M_ItfFlyingSawStateFMData := THIS^;
	ITFFLYINGSAWPROCESSING : L_TS2P_IFlyingSawProcessing := THIS^;
	MASTERVALUES_INT : L_MC1P_IAXIS_REF_MASTERVALUES;
	PDATA : POINTER TO L_TS2M_scData_FM_FlyingSaw;
	PPAR : POINTER TO L_TS2P_scPar_TM_FlyingSawState;
	PAP : POINTER TO L_TS2P_scAP_TM_FlyingSawState;
	PSF : POINTER TO L_TS2P_scSF_TM_FlyingSawState;
	FB_TRANSITION2STOPSAWERROR : L_UBUP_RequestTransitionLevel;
	FB_TRANSITION2STOPSAW : L_UBUP_RequestTransitionLevel;
	FB_TRANSITION2STARTSAW : L_UBUP_RequestTransitionEdge;
	FB_TRANSITION2STARTSAWMODECHANGE : L_UBUP_RequestTransitionEdge;
	FB_TRANSITION2SYNCINSTANT : L_UBUP_RequestTransitionEdge;
	FB_TRANSITION2SYNCLENGTHCTRLAUTO : L_UBUP_RequestTransitionLevel;
	FB_TRANSITION2SYNCLENGTHCTRLRESUME : L_UBUP_RequestTransitionEdge;
	FB_TRANSITION2SYNCMARKCTRL : L_UBUP_RequestTransitionEdge;
	FB_TRANSITION2SYNCMARKCTRLRESUME : L_UBUP_RequestTransitionEdge;
	FB_TRANSITION2SYNCSETCUTLENGTHINST : L_UBUP_RequestTransitionEdge;
	FB_TRANSITION2SYNCAFTERSYNCOUT : L_UBUP_RequestTransitionEdge;
	FB_TRANSITION2SYNCAFTERWAITING : L_UBUP_RequestTransitionLevel;
	FB_TRANSITION2SYNCFROMMOVETOLOWERLIMIT : L_UBUP_RequestTransitionEdge;
	FB_TRANSITION2SYNCFROMSYNCOUT : L_UBUP_RequestTransitionEdge;
	FB_TRANSITION2SYNCNEXTCUT : L_UBUP_RequestTransitionEdge;
	FB_TRANSITION2SYNCRESETMARKSTACK : L_UBUP_RequestTransitionEdge;
	FB_TRANSITION2SYNCOUTNEXTCUT : L_UBUP_RequestTransitionEdge;
	FB_TRANSITION2SYNCOUTRESETMARKSTACK : L_UBUP_RequestTransitionEdge;
	FB_TRANSITION2SAWSYNCHRONIZED : L_UBUP_RequestTransitionEdge;
	FB_TRANSITION2SAWSYNCHRONIZEDAFTERMOVEGAP : L_UBUP_RequestTransitionEdge;
	FB_TRANSITION2MOVETOLOWERLIMIT : L_UBUP_RequestTransitionEdge;
	FB_TRANSITION2WAITINGFORNEXTCUT : L_UBUP_RequestTransitionEdge;
	FB_TRANSITION2MOVEGAP : L_UBUP_RequestTransitionEdge;
	FB_MATERIALCOUNTER : L_TS2P_MaterialCounter;
	FB_CALCULATETARGETPOS : L_TS2P_CalculateTargetPos;
	FB_PROCESSCONTROL : L_TS2P_ProcessControl;
	FB_POSPROFILERCLUTCH : L_MB1P_PosProfilerClutchHigh;
	FB_CONTROLSETVALUES : L_MC1P_ControlSetValues;
	FB_L_TB2P_TP_CONVERTER : L_TB2P_TP_Converter;
	FB_MARKSTACK : L_TS2P_MarkStackFlyingSaw;
	FB_SYNCHRONISEDOVERRIDE : L_TS2P_SyncronisedOverride;
	FB_INPOSITION : L_TT1P_InPosition;
	FB_XEXECUTENEXTCUT_R_TRIG : R_TRIG;
	FB_XRESETMARKSTACK_R_TRIG : R_TRIG;
	XINITDONE : BOOL;
	XEXITDONE : BOOL;
	C_LRMATERIALCOUNTERCYCLELENGTH : LREAL := (16#4FFFFFFFFFFFFFFF * 1E-08);
	FLYINGSAWPROCESSING : L_TS2P_IFlyingSawProcessing;
	FMDATA : L_TS2M_ItfFlyingSawStateFMData;
	GET_LRACTIVEDEC : LREAL;
	GET_LRACTIVEJERK : LREAL;
END_VAR
END_FUNCTION_BLOCK

METHOD CALL_CALCBALANCEDPROFILE
END_METHOD

METHOD CALL_CHECKMASTERNOISE
END_METHOD

METHOD CHECKSYNCHRONISED : BOOL
END_METHOD

METHOD CALLFBS
VAR_INPUT
	ECASE : L_UBUP_StateHandleCase;
END_VAR
END_METHOD

METHOD CALLSTATE
VAR_INPUT
	ITFSTATESERVER : L_UBUP_IStateServer;
	ISTATE : INT;
	ECASE : L_UBUP_StateHandleCase;
END_VAR
END_METHOD

METHOD CHECKTRANSITION
VAR_INPUT
	ITFSTATESERVER : L_UBUP_IStateServer;
END_VAR
END_METHOD

METHOD DISABLECLIENT : BOOL
VAR_INPUT
	XFIRSTCALL : BOOL;
END_VAR
END_METHOD

METHOD ENABLECLIENT : BOOL
VAR_INPUT
	XFIRSTCALL : BOOL;
END_VAR
END_METHOD

METHOD FINALIZECYCLE
END_METHOD

METHOD LEAVESTATE
END_METHOD

METHOD PREPARECYCLE
END_METHOD

METHOD STIMULATETRANSITION
VAR_INPUT
	ECASE : L_UBUP_StateHandleCase;
END_VAR
END_METHOD

METHOD STATE_EXIT : BOOL
VAR_INPUT
	ECASE : L_UBUP_StateHandleCase;
END_VAR
END_METHOD

METHOD FB_INIT : BOOL
VAR_INPUT
	BINITRETAINS : BOOL;
	BINCOPYCODE : BOOL;
END_VAR
END_METHOD

METHOD CALL_ALLOCPOINTADR
END_METHOD

METHOD CALL_EXIT_CALLFBS
END_METHOD

METHOD CALL_MASTERAXISREF
VAR_INPUT
	MASTERVALUES : L_MC1P_IAXIS_REF_MASTERVALUES;
END_VAR
END_METHOD

METHOD CALL_RESETOUTPUT
END_METHOD

METHOD STATE_MOVE_GAP
VAR_INPUT
	ECASE : L_UBUP_StateHandleCase;
	ITFSTATESERVER : L_UBUP_IStateServer;
END_VAR
END_METHOD

METHOD STATE_MOVE_TO_LOWER_LIMIT
VAR_INPUT
	ECASE : L_UBUP_StateHandleCase;
	ITFSTATESERVER : L_UBUP_IStateServer;
END_VAR
END_METHOD

METHOD STATE_SAW_SYNCHRONIZED
VAR_INPUT
	ECASE : L_UBUP_StateHandleCase;
	ITFSTATESERVER : L_UBUP_IStateServer;
END_VAR
END_METHOD

METHOD STATE_SAW_SYNCHRONIZING
VAR_INPUT
	ECASE : L_UBUP_StateHandleCase;
	ITFSTATESERVER : L_UBUP_IStateServer;
END_VAR
END_METHOD

METHOD STATE_START_SAW
VAR_INPUT
	ECASE : L_UBUP_StateHandleCase;
	ITFSTATESERVER : L_UBUP_IStateServer;
END_VAR
END_METHOD

METHOD STATE_STOP_SAW
VAR_INPUT
	ECASE : L_UBUP_StateHandleCase;
	ITFSTATESERVER : L_UBUP_IStateServer;
END_VAR
END_METHOD

METHOD STATE_SYNC_OUT
VAR_INPUT
	ECASE : L_UBUP_StateHandleCase;
	ITFSTATESERVER : L_UBUP_IStateServer;
END_VAR
END_METHOD

METHOD STATE_WAITING_FOR_NEXT_CUT
VAR_INPUT
	ECASE : L_UBUP_StateHandleCase;
	ITFSTATESERVER : L_UBUP_IStateServer;
END_VAR
END_METHOD

METHOD CALL_FB_CALCULATETARGETPOS
END_METHOD

METHOD CALL_FB_CONTROLSETVALUES
END_METHOD

METHOD CALL_FB_INPOSITION
END_METHOD

METHOD CALL_FB_L_TB2P_TP_CONVERTER
END_METHOD

METHOD CALL_FB_MATERIALCOUNTER
END_METHOD

METHOD CALL_FB_PROCESSCONTROL
END_METHOD

METHOD CALL_FB_SYNCHRONISEDOVERRIDE
END_METHOD

METHOD TRANS_TO_SAW_SYNCHRONIZED : BOOL
END_METHOD

METHOD CLUTCH
VAR_INPUT
	ITFTECHMODULE : L_TS2P_IFlyingSawProcessing;
	XENABLE : BOOL;
	XSYNCVEL : BOOL := FALSE;
	XSYNCPOS : BOOL;
	XSYNCOUTINSTANT : BOOL;
	LRSYNCVEL : LREAL := 10;
	LRSYNCACC : LREAL := 100;
	LRSYNCDEC : LREAL := 100;
	LRSYNCJERK : LREAL := 10000;
	LRCYCMASTERPOS : LREAL;
	LRCYCMASTERVEL : LREAL;
	LRCYCMASTERACC : LREAL;
	LRSETSLAVEPOS : LREAL;
	LRSETSLAVEVEL : LREAL;
	LRSETSLAVEACC : LREAL;
END_VAR
VAR_OUTPUT
	EERRORID : L_IE1P.L_IE1P_Error;
	XERROR : BOOL;
	XBUSY : BOOL;
	XDONE : BOOL;
	XACCDECSYNC : BOOL;
	XVELSYNCHRONISED : BOOL;
	XPOSSYNCHRONISED : BOOL;
	LRSETSLAVEPOSOUT : LREAL;
	LRSETSLAVEVELOUT : LREAL;
	LRSETSLAVEACCOUT : LREAL;
	XPROFILERESETTIMEVALID : BOOL;
	LRPROFILERESETTIME : LREAL;
END_VAR
END_METHOD

METHOD EXECUTEGAP
VAR_INPUT
	ITFTECHMODULE : L_TS2P_IFlyingSawProcessing;
	XENABLE : BOOL;
	LRSYNCVEL : LREAL := 10;
	LRSYNCACC : LREAL := 100;
	LRSYNCDEC : LREAL := 100;
	LRSYNCJERK : LREAL := 10000;
	XEXECUTEGAP : BOOL;
	XAUXEXECUTEGAP : BOOL := FALSE;
	LRCYCMASTERPOS : LREAL;
	LRCYCMASTERVEL : LREAL;
	LRCYCMASTERACC : LREAL;
	LRSETSLAVEPOS : LREAL;
	LRSETSLAVEVEL : LREAL;
	LRSETSLAVEACC : LREAL;
END_VAR
VAR_OUTPUT
	EERRORID : L_IE1P.L_IE1P_Error;
	XERROR : BOOL;
	XBUSY : BOOL;
	XDONE : BOOL;
	XACCDECSYNC : BOOL;
	XVELSYNCHRONISED : BOOL;
	XPOSSYNCHRONISED : BOOL;
	LRSETSLAVEPOSOUT : LREAL;
	LRSETSLAVEVELOUT : LREAL;
	LRSETSLAVEACCOUT : LREAL;
	XPROFILERESETTIMEVALID : BOOL;
	LRPROFILERESETTIME : LREAL;
END_VAR
END_METHOD

METHOD MARKSTACK_GETMARK
VAR_INPUT
	ITFTECHMODULE : L_TS2P_IFlyingSawProcessing;
	XENABLE : BOOL;
	XGETMARK : BOOL;
	XRESETGETMARK : BOOL;
	XRESETMARKSTACK : BOOL;
	LRCYCSETPOS : LREAL;
	LRCYCSETVEL : LREAL;
END_VAR
VAR_OUTPUT
	XMARKSTACKFULL : BOOL;
	XMARKSTACKEMPTY : BOOL;
	WMARKSINSTACK : WORD;
	XMARKVALID : BOOL;
	LRMARKPOSOUT : LREAL;
END_VAR
END_METHOD

METHOD MARKSTACK_SETMARK
VAR_INPUT
	ITFTECHMODULE : L_TS2P_IFlyingSawProcessing;
	XENABLE : BOOL;
	XSETMARK : BOOL;
	LRMARKPOS : LREAL;
	XRESETMARKSTACK : BOOL;
	LRCYCSETPOS : LREAL;
	LRCYCSETVEL : LREAL;
END_VAR
VAR_OUTPUT
	XMARKSTACKFULL : BOOL;
	XMARKSTACKEMPTY : BOOL;
	WMARKSINSTACK : WORD;
	XNEWMARKRECEIVED : BOOL;
END_VAR
END_METHOD

METHOD POSITIONING
VAR_INPUT
	ITFTECHMODULE : L_TS2P_IFlyingSawProcessing;
	XENABLE : BOOL;
	XMOVETOTARGETPOS : BOOL;
	LRTARGETPOS : LREAL;
	LRPOSITIONINGVEL : LREAL;
	LRPOSITIONINGACC : LREAL;
	LRPOSITIONINGDEC : LREAL;
	LRPOSITIONINGJERK : LREAL;
	LRSETSLAVEPOS : LREAL;
	LRSETSLAVEVEL : LREAL;
	LRSETSLAVEACC : LREAL;
	LRCORRECTTIMEBASE : LREAL := 0;
	LROVERRIDE : LREAL := 1.0;
END_VAR
VAR_OUTPUT
	EERRORID : L_IE1P.L_IE1P_Error;
	XERROR : BOOL;
	XBUSY : BOOL;
	XDONE : BOOL;
	XPOSITIONING : BOOL;
	XINPOSITION : BOOL;
	LRSETSLAVEPOSOUT : LREAL;
	LRSETSLAVEVELOUT : LREAL;
	LRSETSLAVEACCOUT : LREAL;
	XPROFILERESETTIMEVALID : BOOL;
	LRPROFILERESETTIME : LREAL;
END_VAR
END_METHOD

(* ---- L_TS2M_TM_FLYINGSAWSTATE.fb ---- *)
FUNCTION_BLOCK L_TS2M_TM_FLYINGSAWSTATE EXTENDS L_TB2M_TM_MotionControl
VAR
	TM_FLYINGSAWSTATECONFIG : L_TB2P_ModuleHandlerConfig;
	PSCINPUT : POINTER TO L_TS2P_FlyingSawStateIn;
	PSCOUTPUT : POINTER TO L_TS2P_FlyingSawStateOut;
	PPAR : POINTER TO L_TS2P_scPar_TM_FlyingSawState;
	PSF : POINTER TO L_TS2P_scSF_TM_FlyingSawState;
	PAP : POINTER TO L_TS2P_scAP_TM_FlyingSawState;
	ITFTMDATA : L_TS2M_ItfFlyingSawStateTMData := THIS^;
	PDATA : POINTER TO L_TS2M_scData_FlyingSawState;
	FB_CONDDIRENABLED_SAWINPROCESS : L_UBUP_ConditionInput;
	FB_CONDDIRENABLED_MOVETOPARKPOS : L_UBUP_ConditionInput;
	FB_CONDCOLLECTSAWINPROCESS : L_UBUP_ConditionCollection := STRUCT(aitfCondition := [fb_ConditionOperationEnabled, fb_ConditionLimiter, fb_ConditionAxisHomed, fb_CondDirEnabled_SawInProcess]);
	FB_CONDCOLLECTMOVETOPARKPOS : L_UBUP_ConditionCollection := STRUCT(aitfCondition := [fb_ConditionOperationEnabled, fb_ConditionLimiter, fb_ConditionAxisHomed, fb_CondDirEnabled_MoveToParkPos]);
	FB_TRANSITION2SAWINPROCESS : L_UBUP_RequestTransitionLevel;
	FB_TRANSITION2MOVETOPARKPOS : L_UBUP_RequestTransitionEdge;
	FB_TRANSITION2MOVETOPARKPOSFROMSAWINPROCESS : L_UBUP_RequestTransitionEdge;
	FB_TRANSITION2HALTFROMSAWINPROCESS : L_UBUP_RequestTransitionEdge;
	FB_MOVETOPARKPOS : MC_MoveAbsolute;
	FB_FM_FLYINGSAW : L_TS2M_FM_FlyingSawState := STRUCT(ErrorManager := fb_ErrorManager);
	_ITFSTRUCTPROVIDERFLYINGSAW : L_TS2P_IStructProviderFlyingSaw;
	_SCTPRECEIVEDATA : L_MC1P_TpReceiveData;
	_FB_TPRECDATAPROXYMARKCORR : L_MC1P_TouchProbeRecDataProxy;
	CONNECTOR : __SYSTEM.IQueryInterface;
	FLYINGSAWPROCESSINGEXTENSION : L_TS2P_IFlyingSawProcessing;
	REMAININGTIMEOFPROFILE : LREAL;
	REMAININGTIMEOFPROFILEAVAILABLE : BOOL;
	TMDATA : L_TS2M_ItfFlyingSawStateTMData;
END_VAR
END_FUNCTION_BLOCK

METHOD CALLFBS
VAR_INPUT
	ECASE : L_UBUP_StateHandleCase;
END_VAR
END_METHOD

METHOD CALLSTATE
VAR_INPUT
	ITFSTATESERVER : L_UBUP_IStateServer;
	ISTATE : INT;
	ECASE : L_UBUP_StateHandleCase;
END_VAR
END_METHOD

METHOD CHECKTRANSITION
VAR_INPUT
	ITFSTATESERVER : L_UBUP_IStateServer;
END_VAR
END_METHOD

METHOD FINALIZECYCLE
END_METHOD

METHOD PREPARECYCLE
END_METHOD

METHOD STIMULATETRANSITION
VAR_INPUT
	ECASE : L_UBUP_StateHandleCase;
END_VAR
END_METHOD

METHOD STATE_ABORT
VAR_INPUT
	ECASE : L_UBUP_StateHandleCase;
	ITFSTATESERVER : L_UBUP_IStateServer;
END_VAR
END_METHOD

METHOD STATE_EXIT : BOOL
VAR_INPUT
	ECASE : L_UBUP_StateHandleCase;
END_VAR
END_METHOD

METHOD STATE_HALT
VAR_INPUT
	ECASE : L_UBUP_StateHandleCase;
	ITFSTATESERVER : L_UBUP_IStateServer;
END_VAR
END_METHOD

METHOD STATE_HOMING
VAR_INPUT
	ECASE : L_UBUP_StateHandleCase;
	ITFSTATESERVER : L_UBUP_IStateServer;
END_VAR
END_METHOD

METHOD STATE_MOVE_TO_PARKPOS
VAR_INPUT
	ECASE : L_UBUP_StateHandleCase;
	ITFSTATESERVER : L_UBUP_IStateServer;
END_VAR
END_METHOD

METHOD STATE_SAW_IN_PROCESS
VAR_INPUT
	ECASE : L_UBUP_StateHandleCase;
	ITFSTATESERVER : L_UBUP_IStateServer;
END_VAR
END_METHOD

METHOD STATE_STANDBY
VAR_INPUT
	ECASE : L_UBUP_StateHandleCase;
	ITFSTATESERVER : L_UBUP_IStateServer;
END_VAR
END_METHOD

METHOD CALL_ALLOCPOINTADR
END_METHOD

METHOD CALL_EXIT_CALLFBS
END_METHOD

METHOD CALL_RESETOUTPUT
END_METHOD

METHOD CALL_FM_FLYINGSAW
END_METHOD

METHOD MOVETOPARKPOS : BOOL
VAR_INPUT
	XEXECUTEMOVETOPARKPOS : BOOL;
	LRPARKPOSITION : LREAL := 180;
	EPOSITIONINGDIRECTION : MC_DIRECTION := MC_DIRECTION.mcPositiveDirection;
	LRPOSITIONINGVEL : LREAL := 10;
	LRPOSITIONINGACC : LREAL := 100;
	LRPOSITIONINGDEC : LREAL := 100;
	LRJERK : LREAL := 0;
END_VAR
VAR_OUTPUT
	XBUSY : BOOL;
	XDONE : BOOL;
	XCOMMANDABORTED : BOOL;
END_VAR
VAR_IN_OUT
	AXIS : AXIS_REF;
END_VAR
END_METHOD

(* ---- L_TS2P_ALLOWEDDIRECTION.fb ---- *)
FUNCTION_BLOCK L_TS2P_ALLOWEDDIRECTION
VAR_INPUT
	XENABLE : BOOL;
	XRESETERROR : BOOL;
	ESETVALUEMODE : L_MC1P_SetValueMode := L_MC1P_SetValueMode.Pos;
	LRSETPOSITION : LREAL;
	LRSETVELOCITY : LREAL;
	LRSETACCELERATION : LREAL;
	LRCYCLELENGTH : LREAL;
	ETRAVERSINGRANGE : L_MC1P_TraversingRange := L_MC1P_TraversingRange.Modulo;
	EALLOWEDDIRECTION : L_TB2P_AllowedDirection;
	LRALLOWEDPOSERROR : LREAL;
END_VAR
VAR_OUTPUT
	XENABLED : BOOL;
	LRSETPOSOUT : LREAL;
	LRSETVELOUT : LREAL;
	LRSETACCOUT : LREAL;
	XLIMITATIONACTIVE : BOOL;
	XWARNING : BOOL;
	XERROR : BOOL;
	EERRORID : WORD;
END_VAR
VAR
	XINITDONE : BOOL;
	LRTASKCYCLETIME : LREAL;
	LRSETPOSOUT_REVERSING : LREAL;
	XVELMODE_INT : BOOL;
	LRPOSDIFF : LREAL := 0;
	LRSETPOSDIFFINTEGRATOR : LREAL := 0;
	LRSETPOSITION_INT : LREAL;
	LRSETVELOCITY_INT : LREAL;
	LRCYCLICPOSDIFF : LREAL;
	LRSETPOSITIONOLD : LREAL;
	XMASTERINDISABLEDDIRECTION : BOOL;
	XRESETERROR_OLD : BOOL;
END_VAR
END_FUNCTION_BLOCK

(* ---- L_TS2P_CALCULATETARGETPOS.fb ---- *)
FUNCTION_BLOCK L_TS2P_CALCULATETARGETPOS
VAR_INPUT
	XRESET : BOOL;
	XENABLE : BOOL;
	XEXECUTENEXTCUT : BOOL;
	XEXECUTEFIRSTCUT : BOOL;
	XSETCUTTINGLENGTHINSTANT : BOOL;
	XTPNOTVALID : BOOL;
	XEXECUTEGAP : BOOL;
	XRESUMETARGETPOS : BOOL;
	XSTARTFLYINGSAW : BOOL;
	ETMSTATE : L_TB2P_States;
	XSYNCININSTANT : BOOL;
	XSETMATERIALCOUNTER : BOOL;
	LRMATERIALCOUNTER : LREAL;
	LRDELTAMATERIALPOS : LREAL;
	LRSLAVEPOS : LREAL;
	LRCUTTINGLENGTH : LREAL;
	LRMARKSENSORPOS : LREAL;
	LRGAP : LREAL;
	LRMARKPOSITION : LREAL;
	XLOADTOTALCUTTINGLENGTH : BOOL;
	LRLOADTOTALCUTTINGLENGTH : LREAL;
	XLOADTARGETPOS : BOOL;
	LRLOADTARGETPOS : LREAL;
	EMODE : L_TS2P_FlyingSawMode;
	LRVELINMASTER : LREAL;
	LRACCDIST : LREAL;
	LRACCTIME : LREAL;
	LRTASKCYCLETIME : LREAL;
	XEMPTYSTACK : BOOL;
	XSYNCHRONIZED : BOOL;
	XINPOSITION : BOOL;
END_VAR
VAR_OUTPUT
	XEXECUTEGAPOUT : BOOL;
	LRTARGETPOS : LREAL;
	LRTARGETPOS_OUT : LREAL;
	LRTOTALPRODUCTLENGTH : LREAL;
	XCUTTINGLENGTHVALID : BOOL;
	LRACTIVECUTTINGLENGTH : LREAL;
END_VAR
VAR
	LROFFSET_INT : LREAL;
	XGAPREQUESTED : BOOL;
	LRDELTAMATERIALPOS_INT : LREAL;
	LRTOLERANCE : LREAL;
	LROFFSETOUT_INT : LREAL;
	LRGAPTOTAL_INT : LREAL;
	XSYNCININSTANT_LOCK : BOOL;
	XENABLE_OLD : BOOL;
	XSYNCININSTANT_OLD : BOOL;
	LRMATERIALCOUNTER_OLD : LREAL;
	XEXECUTENEXTCUT_OLD : BOOL;
	XEXECUTEGAP_OLD : BOOL;
	XEXECUTEFIRSTCUT_OLD : BOOL;
	EMODE_OLD : WORD;
	ETMSTATE_OLD : L_TB2P_States;
	XTPNOTVALID_OLD : BOOL;
	XSETCUTTINGLENGTHINSTANT_OLD : BOOL;
	XSETMATERIALCOUNTER_OLD : BOOL;
	LRMARKPOSITION_OLD : LREAL;
END_VAR
END_FUNCTION_BLOCK

(* ---- L_TS2P_CALCULATETPCOMPENSATIONFACTOR.fb ---- *)
FUNCTION_BLOCK L_TS2P_CALCULATETPCOMPENSATIONFACTOR
VAR_OUTPUT
	LRFACTOR : LREAL;
	LRCOMPENSATIONCYCLES : LREAL;
END_VAR
VAR_IN_OUT
	TPAXIS : AXIS_REF;
END_VAR
VAR
	LRSETPOSARRAY : ARRAY [0..15] OF LREAL;
	BYCOUNTER : BYTE;
	LRTEMP : LREAL;
	LRPOSDIFF : LREAL;
	LRSETACTDIFF : LREAL;
	XERRORINVALIDAXIS : BOOL;
	LRSETPOS : LREAL;
	LRACTPOS : LREAL;
	LRCYCLELENGTH : LREAL;
	LRADDITIONALCORRECTION : LREAL;
	LRTEMP2 : LREAL;
	XINCREMENTCYCLES : BOOL;
END_VAR
END_FUNCTION_BLOCK

METHOD SEARCHARRAY
END_METHOD

(* ---- L_TS2P_CALCULATETPONMATERIALPOS.fb ---- *)
FUNCTION_BLOCK L_TS2P_CALCULATETPONMATERIALPOS
VAR_INPUT
	XENABLE : BOOL;
	BYTASKCYCLEDELAY : BYTE := 4;
	XMARKRECEIVE : BOOL;
	LRMARKSENSORPOS : LREAL;
	LRACTMARKPOSIN : LREAL;
	LRCYCPOSTPAXIS : LREAL;
	LRCYCVELTPAXIS : LREAL;
	LRCYCLELENGTHTPAXIS : LREAL;
	LRCYCLELENGTHTARGETAXIS : LREAL;
	LRTASKCYCLETIME : LREAL;
	XRESETMARKSTACK : BOOL;
	LRMATERIALCOUNTER : LREAL;
	LRUPPERLIMITWORKINGRANGE : LREAL;
	LRLOWERLIMITWORKINGRANGE : LREAL;
	LRFACTOR : LREAL;
	LRCOMPVELFACTOR : LREAL;
	XSCIPTONEXTPOSOUT : BOOL;
	XSYNCININSTANT : BOOL;
	XEXECUTEFIRSTCUT : BOOL;
END_VAR
VAR_OUTPUT
	LRTPPOSOUT : LREAL;
	XEXECUTEFIRSTCUT_OLD : BOOL;
	LRTPACTTIMESTAMP : LREAL;
	XFULL : BOOL;
	WMARKPOSITIONVALID : WORD;
	WININDEX : WORD;
	ALRMARKPOSITIONARRAY : ARRAY [0..15] OF LREAL := [0, 0, 0, 0, 0, 0, 0, 0, 0, 0, 0, 0, 0, 0, 0, 0];
	ALRTIMESTAMPARRAY : ARRAY [0..15] OF LREAL;
	XEMPTY : BOOL := TRUE;
	WOUTINDEX : WORD;
	BYREMAINMARKSTACK : BYTE := 15;
	XTPRECEIVED : BOOL;
	XMARKRECEIVED : BOOL;
	XTPPOSVALID : BOOL;
	BYCOUNTEROUT : BYTE;
	XERROR : BOOL;
END_VAR
VAR
	R_TRIG1 : R_TRIG;
	LRTIMESTAMP : LREAL;
	BYTPIDLEINDEX : BYTE;
	BYTPACTINDEX : BYTE;
	ALRPOSITION : ARRAY [0..15] OF LREAL;
	BYTPPREVINDEX : BYTE;
	BYTMP : BYTE;
	XSKIPTONEXTPOS : BOOL;
	WTESTCOUNTER : WORD;
	XTEST : BOOL;
	XWAIT : BOOL;
	WCOUNTINVALIDTIMESTAMP : WORD;
	LRDISTINACTMASTER : LREAL;
	BYTEST : BYTE;
	LRMARKPOSITIONDIFF : LREAL;
	LRMARKPOSITIONDIFF2 : LREAL;
	LRPOSFIFOX : ARRAY [1..20] OF LREAL := [10(0)];
	LRPOSFIFOREG : ARRAY [1..20] OF LREAL := [10(0)];
	BYCOUNTER : BYTE := 1;
	LRSTACKDIFFERENCE : LREAL;
	LRTPDELTAINMS : LREAL;
	LRDELTAPCT : LREAL;
	LRTEMP : LREAL;
	IDIRECTION : INT;
	LRACTMARKPOSIN_OLD : LREAL;
	R_TRIG2 : R_TRIG;
	DWSTATE : DWORD;
	WSTOREDPOSVALUES : WORD;
	LRACTMARKPOSIN_INT : LREAL;
	XSYNCININSTANT_OLD : BOOL;
	XWAIT_OLD : BOOL;
	XRESETMARKSTACK_OLD : BOOL;
	BYCNT : BYTE;
	BYSTEPPER : BYTE;
END_VAR
END_FUNCTION_BLOCK

METHOD SEARCHINSTACKNEGATIVE
END_METHOD

METHOD SEARCHINSTACKPOSITIVE
END_METHOD

(* ---- L_TS2P_CAMCREATOR.fb ---- *)
FUNCTION_BLOCK L_TS2P_CAMCREATOR
VAR_INPUT
	XENABLEINTERNALCAMTABLE : BOOL;
	XEXECUTE : BOOL;
	PCAMPOINTS : POINTER TO L_MC2P_CamDataXYVA;
	INUMOFPOINTS : INT;
	LRMASTERMAXVEL : LREAL;
	LRMASTERMAXACC : LREAL;
	LRMASTERSCALING : LREAL := 1;
	LRSLAVESCALING : LREAL := 1;
END_VAR
VAR_OUTPUT
	XINTERNALCAMTABLELACTIVE : BOOL;
	XERROR : BOOL;
	EERRORID : L_IE1P_Error;
	XBUSY : BOOL;
	XDONE : BOOL;
	CAMTABLEOUT : MC_CAM_REF;
	LRSLAVEMAXPOS : LREAL;
	LRSLAVEMINPOS : LREAL;
	LRSLAVEMAXVEL : LREAL;
	LRSLAVEMINVEL : LREAL;
	LRSLAVEMAXACC : LREAL;
	LRSLAVEMINACC : LREAL;
END_VAR
VAR_IN_OUT
	SLAVE : AXIS_REF;
END_VAR
VAR
	EFMSTATE : L_MB1P_States := L_MB1P_States.INIT;
	SMC_CAMBOUNDS1 : L_MC2P_BoundsCam;
	SMC_CAMBOUNDSINIT : L_MC2P_BoundsCam;
	CAMREF : L_MC2P_CamRefFromStruct;
	PCAMPOINTS_INT : POINTER TO L_MC2P_CamDataXYVA;
	INUMOFPOINTS_INT : INT;
	XINTERNALCONTROL : BOOL;
	XEXECUTE_OLD : BOOL;
	ASCCAMPOINTS : ARRAY [0..30] OF L_MC2P_CamDataXYVA;
	XINVALIDCAMTABLE : BOOL;
	XVISUACTIVE : BOOL := TRUE;
	DIFRAME : DINT;
	DIFRAME_OLD : DINT;
	ARVISPOINTLINES : ARRAY [1..10] OF L_MC2P_CamDataXYVA;
	IVISUTABLESETPOS : INT := 0;
	IVISUTABLESETPOS_OLD : INT := 0;
	IVISUTABLEMAXPOS : INT := 30;
	IVISSHOWLINESNO : INT;
	XVISPOINTMIN : BOOL;
	XVISPOINTMAX : BOOL;
	XVISUSETPOSUP : BOOL;
	XVISUSETPOSDOWN : BOOL;
	XVISUSETPOSUP_OLD : BOOL;
	XVISUSETPOSDOWN_OLD : BOOL;
	XSCROLBUTTENACTIVE : BOOL;
	TSETTIME : TIME := TIME#400ms;
	TON_SCROLBUTTEN : TON;
END_VAR
END_FUNCTION_BLOCK

METHOD CALL_CAMBOUNDS
VAR_IN_OUT
	SLAVE : AXIS_REF;
END_VAR
END_METHOD

METHOD CALL_CAMREF
END_METHOD

METHOD CALL_CAMTABLEEQUIDISTANT
END_METHOD

METHOD CALL_CAMTABLENONEQUIDISTANT
END_METHOD

METHOD CALL_CAMTABLEPOLYNOMIAL
END_METHOD

METHOD CALL_ERRORHANDLER
END_METHOD

METHOD CALL_FBMETHODS
VAR_IN_OUT
	SLAVE : AXIS_REF;
END_VAR
END_METHOD

METHOD CALL_INTERNALCTRL
END_METHOD

METHOD CALL_OUTPUT
END_METHOD

METHOD CALL_RESETCOMMANDS
VAR_IN_OUT
	SLAVE : AXIS_REF;
END_VAR
END_METHOD

METHOD CALL_RESETOUTPUT
END_METHOD

METHOD CALL_STATEMACHINE
END_METHOD

METHOD CALL_VIS_TON_SCROLBUTTEN
END_METHOD

METHOD CALL_VISUTABCTRL
END_METHOD

METHOD CALL_VISUUPDATETAB
END_METHOD

METHOD DISABALE_VISU
END_METHOD

METHOD ENABLE_VISU
END_METHOD

METHOD CALL_S000_CYCLIC
END_METHOD

METHOD CALL_S001_INIT
END_METHOD

METHOD CALL_S002_READY
END_METHOD

(* ---- L_TS2P_CAMTABLEINFO.fb ---- *)
FUNCTION_BLOCK L_TS2P_CAMTABLEINFO
VAR_INPUT
	XENABLE : BOOL;
	CAMTABLE : MC_CAM_REF;
	LRMASTERMAXVEL : LREAL := 100;
	LRMASTERMAXACC : LREAL := 1000;
	LRMASTERSCALING : LREAL := 1;
	LRSLAVESCALING : LREAL := 1;
END_VAR
VAR_OUTPUT
	XBUSY : BOOL;
	XDONE : BOOL;
	XCAMTABLEVALID : BOOL;
	LRMASTERSTARTPOS : LREAL;
	LRMASTERENDPOS : LREAL;
	LRSLAVESTARTPOS : LREAL;
	LRSLAVEENDPOS : LREAL;
	LRSLAVEMAXPOS : LREAL;
	LRSLAVEMINPOS : LREAL;
	LRSLAVEMAXVEL : LREAL;
	LRSLAVEMINVEL : LREAL;
	LRSLAVEMAXACC : LREAL;
	LRSLAVEMINACC : LREAL;
END_VAR
VAR_IN_OUT
	SLAVEAXIS : AXIS_REF;
END_VAR
VAR
	ESTATE : L_MB1P_States := L_MB1P_States.INIT;
	CAMTABLE_INT : MC_CAM_REF;
	PCAMDATA_INT : POINTER TO L_MC2P_CamData;
	LRMASTERMAXVEL_INT : LREAL := 0;
	LRMASTERMAXACC_INT : LREAL := 0;
	LRMASTERSCALING_INT : LREAL := 0;
	LRSLAVESCALING_INT : LREAL := 0;
	XENABLE_OLD : BOOL;
	SMC_CAMBOUNDS1 : L_MC2P_BoundsCam;
	XCALCNEWVALUES : BOOL;
END_VAR
END_FUNCTION_BLOCK

METHOD CALC_STARTENDVALUES
END_METHOD

METHOD CALL_CAMBOUNDS
END_METHOD

METHOD CALL_FBMETHODS
END_METHOD

METHOD CALL_OUTPUT
END_METHOD

METHOD CALL_RESETCOMMANDS
END_METHOD

METHOD CALL_RESETOUTPUT
END_METHOD

METHOD CALL_STATEMACHINE
END_METHOD

METHOD GET_XCALCNEWVALUES : BOOL
END_METHOD

METHOD GET_XCRITICALCYCLE : BOOL
END_METHOD

(* ---- L_TS2P_CONDITIONLIMITERSYNCIN.fb ---- *)
FUNCTION_BLOCK L_TS2P_CONDITIONLIMITERSYNCIN EXTENDS L_UBUP_ConditionBase
VAR_INPUT
	ESYNCDIRECTION : L_TS2P_SyncDirection;
	DWLIMITERCONTROL : DWORD;
END_VAR
VAR_OUTPUT
	XDIRECTIONDISABLED : BOOL;
	XINVALIDINPUT : BOOL;
END_VAR
VAR_IN_OUT
	AXIS : AXIS_REF;
END_VAR
END_FUNCTION_BLOCK

METHOD VERIFY : BOOL
VAR_OUTPUT
	XCONDITIONERROR : BOOL;
	EERRORIDPROPOSED : L_IE1P.L_IE1P_Error;
END_VAR
END_METHOD

(* ---- L_TS2P_CONDITIONLOCKTOCAM.fb ---- *)
FUNCTION_BLOCK L_TS2P_CONDITIONLOCKTOCAM EXTENDS L_UBUP_ConditionBase
VAR_IN_OUT
	SCPAR : L_TS2P_scPar_TM_FlexCam;
END_VAR
END_FUNCTION_BLOCK

METHOD VERIFY : BOOL
VAR_OUTPUT
	XCONDITIONERROR : BOOL;
	EERRORIDPROPOSED : L_IE1P.L_IE1P_Error;
END_VAR
END_METHOD

(* ---- L_TS2P_CONDITIONSYNCPARAMETER.fb ---- *)
FUNCTION_BLOCK L_TS2P_CONDITIONSYNCPARAMETER EXTENDS L_UBUP_ConditionBase
VAR_IN_OUT
	SCPAR : L_TS2P_scPar_TM_SyncPosBase;
END_VAR
END_FUNCTION_BLOCK

METHOD VERIFY : BOOL
VAR_OUTPUT
	XCONDITIONERROR : BOOL;
	EERRORIDPROPOSED : L_IE1P.L_IE1P_Error;
END_VAR
END_METHOD

(* ---- L_TS2P_CONDITIONVALIDCAMTABLE.fb ---- *)
FUNCTION_BLOCK L_TS2P_CONDITIONVALIDCAMTABLE EXTENDS L_UBUP_ConditionBase
VAR_INPUT
	WSETCAMTABLE : WORD;
	CAMTABLE1 : MC_CAM_REF;
	CAMTABLE2 : MC_CAM_REF;
	CAMTABLE3 : MC_CAM_REF;
	CAMTABLE4 : MC_CAM_REF;
END_VAR
END_FUNCTION_BLOCK

METHOD VERIFY : BOOL
VAR_OUTPUT
	XCONDITIONERROR : BOOL;
	EERRORIDPROPOSED : L_IE1P.L_IE1P_Error;
END_VAR
END_METHOD

(* ---- L_TS2P_CROSSCUTTERSTATE.fb ---- *)
FUNCTION_BLOCK L_TS2P_CROSSCUTTERSTATE EXTENDS L_TB2P_TechModuleBase
VAR_INPUT
	XENABLE : BOOL;
	XENABLEOPERATION : BOOL;
	XRESETERROR : BOOL;
	XQSPAPPLICATION : BOOL;
	XABORT : BOOL;
	XJOGPOS : BOOL;
	XJOGNEG : BOOL;
	XHOMEEXECUTE : BOOL;
	LROVERRIDE : LREAL := 1;
	SCCTRLBASICMOTION : L_TB2P_scCtrlBasicMotion;
	SCPAR : L_TS2P_scPar_CrossCutterState;
	SCACCESSPOINTS : L_TS2P_scAP_CrossCutterState;
	MASTERVALUES : L_MC1P_IAXIS_REF_MASTERVALUES;
	XEXECUTEMOVETOPARKPOS : BOOL;
	XSYNCIN : BOOL;
	XHOLDINPARKPOS : BOOL;
	LRPRODUCTLENGTH : LREAL;
	LROVERSPEED : LREAL;
	LRSETOFFSETPOSX : LREAL;
	XTRIMPOS : BOOL;
	XTRIMNEG : BOOL;
	XTRIMRESET : BOOL;
	SCTPRECDATA_MARKSENSOR : L_MC1P_TpReceiveData;
	SCTPRECDATA_TOOLSENSOR : L_MC1P_TpReceiveData;
	XTEACHMARKWINDOW : BOOL;
	XTEACHMARKWINDOWTOOL : BOOL;
	XGEARFACTORCORR : BOOL;
	XGEARFACTORCORRHOLD : BOOL;
END_VAR
VAR_OUTPUT
	XREADYFOROPERATION : BOOL;
	XOPERATIONENABLED : BOOL;
	XREADYFORMOTION : BOOL;
	XERROR : BOOL;
	XWARNING : BOOL;
	EERRORID : L_IE1P_Error;
	XSTOACTIVE : BOOL;
	XQSPACTIVE : BOOL;
	XABORTBUSY : BOOL;
	XABORTDONE : BOOL;
	XJOGGINGBUSY : BOOL;
	XHOMINGBUSY : BOOL;
	XHOMINGDONE : BOOL;
	XISHOMED : BOOL;
	ETMSTATE : L_TB2P_States;
	SCSTATUSBASICMOTION : L_TB2P_scStatusBasicMotion;
	LRACTVEL : LREAL;
	LRSETVELOUT : LREAL;
	LRACTPOS : LREAL;
	LRSETPOSOUT : LREAL;
	LRACTFOLLOWINGERROR : LREAL;
	SCSIGNALFLOW : L_TS2P_scSF_CrossCutterState;
	XSYNCHRONISED : BOOL;
	XACCDECSYNC : BOOL;
	XOFFSETTRIMACTIVE : BOOL;
	XINPARKPOS : BOOL;
	XHOLDINPARKPOSACTIVE : BOOL;
	XCUTDONE : BOOL;
	XCUTTINGACTIVE : BOOL;
	LRACTCUTLENGTH : LREAL;
	LROFFSETTOTAL : LREAL;
	XTRQCTRLACTIVE : BOOL;
	LRSETMARKCORROUT : LREAL;
	XMARKWINDOWTEACHED : BOOL;
	LRGEARFACTORCORR : LREAL;
	LRSETTOOLCORROUT : LREAL;
	XMARKWINDOWTEACHEDTOOL : BOOL;
END_VAR
VAR_IN_OUT
	AXIS : AXIS_REF;
END_VAR
VAR
	TM_INT : L_TS2P_TM_CrossCutterState := STRUCT(ModuleHandler := ModuleHandler);
	SCPAR_INT : L_TS2P_scPar_CrossCutterState;
	_UICALLMFUNIDXINPUT : UINT := 1;
	_UICALLMFUNIDXOUTPUT : UINT := 1;
	_MCCALL : L_UM1P_MCCall;
	_ASCINPUT : ARRAY [1.._MCCall.c_BufferDepthInput] OF L_TS2P_CrossCutterStateIn;
	_ASCOUTPUT : ARRAY [1.._MCCall.c_BufferDepthOutput] OF L_TS2P_CrossCutterStateOut;
	_ASCPARCORE : ARRAY [1.._MCCall.c_BufferDepthInput] OF L_TS2P_scPar_CrossCutterState;
	_ASCACCESSPOINTSCORE : ARRAY [1.._MCCall.c_BufferDepthInput] OF L_TS2P_scAP_CrossCutterState;
	_ASCSIGNALFLOWCORE : ARRAY [1.._MCCall.c_BufferDepthOutput] OF L_TS2P_scSF_CrossCutterState;
	_SCINPUTVISU : L_TS2P_CrossCutterStateIn;
	_PSCINPUTVISU : POINTER TO L_TS2P_CrossCutterStateIn := ADR(_scInputVisu);
	_PSCOUTPUTVISU : POINTER TO L_TS2P_CrossCutterStateOut := ADR(_ascOutput[1]);
	_PSCPARVISU : POINTER TO L_TS2P_scPar_CrossCutterState := ADR(scPar_int);
	ITFITECHMODULEINTERNAL : L_TB2P_ITechModuleInternal;
	LRJERKDEC : LREAL;
	LRJOGGINGJERKDEC : LREAL;
	REMAININGTIMEOFPROFILE : LREAL;
	REMAININGTIMEOFPROFILEAVAILABLE : BOOL;
END_VAR
END_FUNCTION_BLOCK

METHOD GET_PAP : POINTER TO L_TB2P_scAP_TM_MotionControl
END_METHOD

METHOD GET_PPAR : POINTER TO L_TB2P_scPar_TM_MotionControl
END_METHOD

METHOD GET_PSF : POINTER TO L_TB2P_scSF_TM_MotionControl
END_METHOD

METHOD CALLFUNCTION
VAR_INPUT
	UIINPUTDATAIDX : UINT;
	UIOUTPUTDATAIDX : UINT;
END_VAR
END_METHOD

METHOD COPYINPUTS : BOOL
VAR_INPUT
	IDX : WORD;
END_VAR
END_METHOD

METHOD COPYOUTPUTS : BOOL
VAR_INPUT
	IDX : WORD;
END_VAR
END_METHOD

METHOD FUNCTIONWASCALLEDTWICE : BOOL
VAR_INPUT
	IDX : WORD;
END_VAR
END_METHOD

METHOD HANDLESTANDARDCALL : BOOL
END_METHOD

METHOD SYNCOUTPUTS
VAR_INPUT
	UICOPYOUTPUTFROMIDX : UINT;
	UICOPYOUTPUTTOIDX : UINT;
END_VAR
END_METHOD

METHOD CALL_INTERNALCTRL
END_METHOD

(* ---- L_TS2P_DISTCORRECTIONWINDOW.fb ---- *)
FUNCTION_BLOCK L_TS2P_DISTCORRECTIONWINDOW
VAR_INPUT
	XENABLE : BOOL;
	XENABLEPOSITION : BOOL;
	LRCYCSETPOSMASTER : LREAL;
	LRCYCLELENGTHMASTER : LREAL;
	LRCYCSETVEL : LREAL;
	XLOADSTARTPOS : BOOL;
	LRSTARTPOS : LREAL;
	XTPRECEIVEDIN : BOOL;
	LRSETCORRECTION : LREAL;
	XCORRWINDOWINXUNITS : BOOL;
	LRSETUPPERWINDOW : LREAL;
	LRSETLOWERWINDOW : LREAL;
	LRCYCPOSFEEDBACK : LREAL;
	DNSETNUMERATORAXISY : DWORD := 1;
	DNSETDENOMINATORAXISY : DWORD := 1;
	LRSETCYCLELENGTHX : LREAL;
	LRSETCYCLELENGTHY : LREAL;
END_VAR
VAR_OUTPUT
	XBUSY : BOOL;
	XCORRECTIONBUSY : BOOL;
	LRSETPOSOUT : LREAL;
	LRSETINTEGRATEDPOSITION : LREAL;
	LRSETPOSCORROUT : LREAL;
	LRSETPOSCORRRESIDUALOUT : LREAL;
	LRDELTAPOSCORROUT : LREAL;
	XCORRNEXTCYCLE : BOOL;
	XERROR : BOOL;
	EERRORID : L_IE1P_Error;
END_VAR
VAR
	LRDELTAPOSTOTAL : LREAL;
	LRMASTERDISTANCE : LREAL;
	LRPOSITIONSET : LREAL;
	LRPOSITIONNORMED : LREAL;
	LRPOSITIONOUTNORMED : LREAL;
	LRDELTAPOSCORRECTION : LREAL;
	LRPOSITIONSETOLD : LREAL;
	LRPOSITIONSETAXISOUT : LREAL;
	BYSTEPPER : BYTE;
	LRCORRECTIONDISTANCELOCAL : LREAL;
	LRCORRECTIONLOCAL : LREAL;
	L_DIFFERENTIATE : L_MC2P_Differentiate;
	INTEGRATOR : L_MC1P_IntegrateAxis;
	LRDELTAPOSOUT : LREAL;
	XEXECUTECORRECTIONINTERN : BOOL;
	XPOSITIVEDIRECTION : BOOL := FALSE;
	LRCORRECTIONDISTANCE : LREAL;
	LRUPPERWINDOWINTERNAL : LREAL;
	LRLOWERWINDOWINTERNAL : LREAL;
	LRTASKCYCLE : LREAL;
	XCORRECTIONACTIVE : BOOL;
	LRCORRECTIONLOCAL1 : LREAL;
	XTPRECEIVEDOLD : BOOL;
	LRINTEGRATORSPEED : LREAL;
	XWINDOWINCYCLE : BOOL;
	LRDELTAWINDOW : LREAL;
	LRCYCPOSINTOOLINTERNAL : LREAL;
	LRUPPERWINDOWINTERNALDELTA : LREAL;
	LRLOWERWINDOWINTERNALDELTA : LREAL;
	XINIT : BOOL := TRUE;
	XINITOUTOFCORRWINDOW : BOOL := TRUE;
	LRLOWERWINDOWINTERNALOLD : LREAL;
	LRUPPERWINDOWINTERNALOLD : LREAL;
	LRCYCPOSFEEDBACKINT : LREAL;
	XCORRECTIONBUSYOLD : BOOL;
	LRSETPOSCORROUTOLD : LREAL;
	LRCYCPOSINTOOLINTERNAL_CASE : LREAL;
	XWINDOWCHANGEDFLAG : BOOL := FALSE;
	LRCYCLELENGTH_INT : LREAL;
	LROFFSET_INT : LREAL;
	LRCYCPOSINTOOLINTERNAL_0LD : LREAL;
	LRPOSITIONNORMED_OLD : LREAL;
	LRPOSITIONNORMED_DIF : LREAL;
	XPOSCORR : BOOL;
	XTPSTORED_INT : BOOL;
	LRSETCORRECTIONSTORED_INT : LREAL;
	XINCORRWINDOW : BOOL;
	XINCORRWINDOWOLD : BOOL;
	LRSETPOSOUTCOMP : LREAL;
	LRCYCPOSINTOOLINTERNALOLD : LREAL;
	LRDELTAPOSOUTINTERNAL : LREAL;
	BYSTEPPEROLD : BYTE := 0;
	LRCYCSETPOSOLD : LREAL;
	LRCORRECTIONINYUNITS : LREAL;
	LRCORRECTIONDISTANCETEMP : LREAL;
END_VAR
END_FUNCTION_BLOCK

METHOD CALL_INIT
END_METHOD

(* ---- L_TS2P_ELECTRONICGEARBOXBASE.fb ---- *)
FUNCTION_BLOCK L_TS2P_ELECTRONICGEARBOXBASE EXTENDS L_TB2P_TechModuleBase
VAR_INPUT
	XENABLE : BOOL;
	XENABLEOPERATION : BOOL;
	XRESETERROR : BOOL;
	XQSPAPPLICATION : BOOL;
	XABORT : BOOL;
	XJOGPOS : BOOL;
	XJOGNEG : BOOL;
	XHOMEEXECUTE : BOOL;
	LROVERRIDE : LREAL := 1;
	SCCTRLBASICMOTION : L_TB2P_scCtrlBasicMotion;
	SCPAR : L_TS2P_scPar_ElectronicGearboxBase;
	SCACCESSPOINTS : L_TS2P_scAP_ElectronicGearboxBase;
	MASTERVALUES : L_MC1P_IAXIS_REF_MASTERVALUES;
	XSYNCIN : BOOL;
	LRSETBASEVEL : LREAL;
	LRSETOFFSETPOS : LREAL;
	LRSETOFFSETVEL : LREAL;
	XTRIMPOS : BOOL;
	XTRIMNEG : BOOL;
	XTRIMRESET : BOOL;
	XINVERTGEARFACTOR : BOOL;
END_VAR
VAR_OUTPUT
	XREADYFOROPERATION : BOOL;
	XOPERATIONENABLED : BOOL;
	XREADYFORMOTION : BOOL;
	XERROR : BOOL;
	XWARNING : BOOL;
	EERRORID : L_IE1P_Error;
	XSTOACTIVE : BOOL;
	XQSPACTIVE : BOOL;
	XABORTBUSY : BOOL;
	XABORTDONE : BOOL;
	XJOGGINGBUSY : BOOL;
	XHOMINGBUSY : BOOL;
	XHOMINGDONE : BOOL;
	XISHOMED : BOOL;
	ETMSTATE : L_TB2P_States := L_TB2P_States.DISABLED;
	SCSTATUSBASICMOTION : L_TB2P_scStatusBasicMotion;
	LRACTVEL : LREAL;
	LRSETVELOUT : LREAL;
	LRACTPOS : LREAL;
	LRSETPOSOUT : LREAL;
	LRACTFOLLOWINGERROR : LREAL;
	SCSIGNALFLOW : L_TS2P_scSF_ElectronicGearboxBase;
	XSYNCHRONISED : BOOL;
	XACCDECSYNC : BOOL;
	XOFFSETTRIMACTIVE : BOOL;
	XBASEVELOCITYACTIVE : BOOL;
	LROFFSETTOTALVEL : LREAL;
END_VAR
VAR_IN_OUT
	AXIS : AXIS_REF;
END_VAR
VAR
	TM_INT : L_TS2P_TM_ElectronicGearboxBase := STRUCT(ModuleHandler := ModuleHandler);
	SCPAR_INT : L_TS2P_scPar_ElectronicGearboxBase;
	_UICALLMFUNIDXINPUT : UINT := 1;
	_UICALLMFUNIDXOUTPUT : UINT := 1;
	_MCCALL : L_UM1P_MCCall;
	_ASCINPUT : ARRAY [1.._MCCall.c_BufferDepthInput] OF L_TS2P_ElectronicGearboxBaseIn;
	_ASCOUTPUT : ARRAY [1.._MCCall.c_BufferDepthOutput] OF L_TS2P_ElectronicGearboxBaseOut;
	_ASCPARCORE : ARRAY [1.._MCCall.c_BufferDepthInput] OF L_TS2P_scPar_ElectronicGearboxBase;
	_ASCACCESSPOINTSCORE : ARRAY [1.._MCCall.c_BufferDepthInput] OF L_TS2P_scAP_ElectronicGearboxBase;
	_ASCSIGNALFLOWCORE : ARRAY [1.._MCCall.c_BufferDepthOutput] OF L_TS2P_scSF_ElectronicGearboxBase;
	_SCINPUTVISU : L_TS2P_ElectronicGearboxBaseIn;
	_PSCINPUTVISU : POINTER TO L_TS2P_ElectronicGearboxBaseIn := ADR(_scInputVisu);
	_PSCOUTPUTVISU : POINTER TO L_TS2P_ElectronicGearboxBaseOut := ADR(_ascOutput[1]);
	_PSCPARVISU : POINTER TO L_TS2P_scPar_ElectronicGearboxBase := ADR(scPar_int);
	ITFITECHMODULEINTERNAL : L_TB2P_ITechModuleInternal;
	LRJERKDEC : LREAL;
	LRJOGGINGJERKDEC : LREAL;
	REMAININGTIMEOFPROFILE : LREAL;
	REMAININGTIMEOFPROFILEAVAILABLE : BOOL;
END_VAR
END_FUNCTION_BLOCK

METHOD GET_PAP : POINTER TO L_TB2P_scAP_TM_MotionControl
END_METHOD

METHOD GET_PPAR : POINTER TO L_TB2P_scPar_TM_MotionControl
END_METHOD

METHOD GET_PSF : POINTER TO L_TB2P_scSF_TM_MotionControl
END_METHOD

METHOD CALLFUNCTION
VAR_INPUT
	UIINPUTDATAIDX : UINT;
	UIOUTPUTDATAIDX : UINT;
END_VAR
END_METHOD

METHOD COPYINPUTS : BOOL
VAR_INPUT
	IDX : WORD;
END_VAR
END_METHOD

METHOD COPYOUTPUTS : BOOL
VAR_INPUT
	IDX : WORD;
END_VAR
END_METHOD

METHOD FUNCTIONWASCALLEDTWICE : BOOL
VAR_INPUT
	IDX : WORD;
END_VAR
END_METHOD

METHOD HANDLESTANDARDCALL : BOOL
END_METHOD

METHOD SYNCOUTPUTS
VAR_INPUT
	UICOPYOUTPUTFROMIDX : UINT;
	UICOPYOUTPUTTOIDX : UINT;
END_VAR
END_METHOD

METHOD CALL_INTERNALCTRL
END_METHOD

(* ---- L_TS2P_FLEXCAMHIGH.fb ---- *)
FUNCTION_BLOCK L_TS2P_FLEXCAMHIGH EXTENDS L_TB2P_TechModuleBase
VAR_INPUT
	XUSEORIGINAL : BOOL;
	XENABLE : BOOL;
	XENABLEOPERATION : BOOL;
	XRESETERROR : BOOL;
	XQSPAPPLICATION : BOOL;
	XABORT : BOOL;
	XJOGPOS : BOOL;
	XJOGNEG : BOOL;
	XHOMEEXECUTE : BOOL;
	LROVERRIDE : LREAL := 1;
	SCCTRLBASICMOTION : L_TB2P_scCtrlBasicMotion;
	SCPAR : L_TS2P_scPar_FlexCamHigh;
	SCACCESSPOINTS : L_TS2P_scAP_FlexCamHigh;
	MASTERVALUES : L_MC1P_IAXIS_REF_MASTERVALUES;
	XCLUTCHCLOSE : BOOL;
	XLOADCLUTCHPOS : BOOL;
	LRLOADCLUTCHPOS : LREAL;
	XFINDCLUTCHXPOS : BOOL;
	XSYNCIN : BOOL;
	XSYNCPOSRESTORE : BOOL;
	XCAMCHANGEINSTANT : BOOL;
	LRSETOFFSETPOSX : LREAL;
	LRSETOFFSETPOSY : LREAL;
	LRSETSCALINGX : LREAL := 1;
	LRSETSCALINGY : LREAL := 1;
	CAMTABLE1 : MC_CAM_REF;
	CAMTABLE2 : MC_CAM_REF;
	CAMTABLE3 : MC_CAM_REF;
	CAMTABLE4 : MC_CAM_REF;
	WSETCAMTABLE : WORD := 1;
	XCAMSEQUENCER : BOOL;
END_VAR
VAR_OUTPUT
	XREADYFOROPERATION : BOOL;
	XOPERATIONENABLED : BOOL;
	XREADYFORMOTION : BOOL;
	XERROR : BOOL;
	XWARNING : BOOL;
	EERRORID : L_IE1P_Error;
	XSTOACTIVE : BOOL;
	XQSPACTIVE : BOOL;
	XABORTBUSY : BOOL;
	XABORTDONE : BOOL;
	XJOGGINGBUSY : BOOL;
	XHOMINGBUSY : BOOL;
	XHOMINGDONE : BOOL;
	XISHOMED : BOOL;
	ETMSTATE : L_TB2P_States;
	SCSTATUSBASICMOTION : L_TB2P_scStatusBasicMotion;
	LRACTVEL : LREAL;
	LRSETVELOUT : LREAL;
	LRACTPOS : LREAL;
	LRSETPOSOUT : LREAL;
	LRACTFOLLOWINGERROR : LREAL;
	SCSIGNALFLOW : L_TS2P_scSF_FlexCamHigh;
	XCLUTCHACTIVE : BOOL;
	XCLUTCHCLOSED : BOOL;
	XACCDECSYNC : BOOL;
	XSYNCHRONISED : BOOL;
	XMOVETOPARKPOSACTIVE : BOOL;
	XINPARKPOS : BOOL;
	XENDOFPROFILE : BOOL;
	LROFFSETPOSX : LREAL;
	LROFFSETPOSY : LREAL;
	LROFFSETSYNCPOS : LREAL;
	WACTIVECAMTABLE : WORD;
	XCAMSEQUENCERACTIVE : BOOL;
END_VAR
VAR_IN_OUT
	AXIS : AXIS_REF;
END_VAR
VAR
	XINTERNALCONTROLACTIVE_OLD : BOOL;
	ITFCONNECTORFLEXCAM : L_TS2P_IConnectorFlexCam;
	TM_INT : L_TS2P_TM_FlexCam;
	SCPAR_INT : L_TS2P_scPar_FlexCamHigh;
	SCDATA_INT : L_TS2P_scData_TM_FlexCam;
	SCDATASP_INT : L_TS2P_scData_TM_FlexCam;
	XUSEORIGINAL_OLD : BOOL;
	_UICALLMFUNIDXINPUT : UINT := 1;
	_UICALLMFUNIDXOUTPUT : UINT := 1;
	_MCCALL : L_UM1P_MCCall;
	_ASCINPUT : ARRAY [1.._MCCall.c_BufferDepthInput] OF L_TS2P_FlexCamHighIn;
	_ASCOUTPUT : ARRAY [1.._MCCall.c_BufferDepthOutput] OF L_TS2P_FlexCamHighOut;
	_ASCPARCORE : ARRAY [1.._MCCall.c_BufferDepthInput] OF L_TS2P_scPar_FlexCamHigh;
	_ASCACCESSPOINTSCORE : ARRAY [1.._MCCall.c_BufferDepthInput] OF L_TS2P_scAP_FlexCamHigh;
	_ASCSIGNALFLOWCORE : ARRAY [1.._MCCall.c_BufferDepthOutput] OF L_TS2P_scSF_FlexCamHigh;
	_SCINPUTVISU : L_TS2P_FlexCamHighIn;
	_PSCINPUTVISU : POINTER TO L_TS2P_FlexCamHighIn := ADR(_scInputVisu);
	_PSCOUTPUTVISU : POINTER TO L_TS2P_FlexCamHighOut := ADR(_ascOutput[1]);
	_PSCDATAVISU : POINTER TO L_TS2P_scData_TM_FlexCam := ADR(scData_int);
	_PSCPARVISU : POINTER TO L_TS2P_scPar_FlexCamHigh := ADR(scPar_int);
	_PSCAPVISU : POINTER TO L_TS2P_scAP_FlexCamHigh;
	_PSCSFVISU : POINTER TO L_TS2P_scSF_FlexCamHigh;
	ITFBASICMOTIONBASE : L_TB2P.L_TB2P_IBasicMotionBase;
	ITFFLEXCAMEXTENSION : L_TS2P_IFlexCam;
	ITFITECHMODULEINTERNAL : L_TB2P_ITechModuleInternal;
	LRJERKDEC : LREAL;
	LRJOGGINGJERKDEC : LREAL;
	REMAININGTIMEOFPROFILE : LREAL;
	REMAININGTIMEOFPROFILEAVAILABLE : BOOL;
END_VAR
END_FUNCTION_BLOCK

METHOD CALL_ABC
VAR_INPUT
	ITFTECHMODULE : L_TB2P.L_TB2P_IBasicMotionBase;
	XQSPAPPLICATION : BOOL;
	XHALT : BOOL;
	XABORT : BOOL;
	XHOMEEXECUTE : BOOL;
	XJOGPOS : BOOL;
	XJOGNEG : BOOL;
	XFINISHPOSITIONING : BOOL;
	XMOVEVELEXECUTE : BOOL;
	XMOVEABSEXECUTE : BOOL;
	XMOVERELEXECUTE : BOOL;
	XENABLEOPERATION : BOOL;
	XRESETERROR : BOOL;
	XENABLEPOSITIVE : BOOL;
	XENABLENEGATIVE : BOOL;
	XDISABLESWLIMIT : BOOL;
	LROVERRIDE : LREAL;
	LROVERRIDEACC : LREAL;
	LROVERRIDEJERK : LREAL;
	XRESETHOMEPOSITION : BOOL;
	XCONTINUOUSUPDATE : BOOL;
	LRPOS_DIST : LREAL;
	LRVEL : LREAL;
	LRACC : LREAL;
	LRDEC : LREAL;
	LRJERK : LREAL;
	EDIRECTION : L_TB2P.MC_DIRECTION;
	SCHOMEEXTTP : L_TB2P.MC_TRIGGER_REF;
	XHOMEABSSWITCH : BOOL;
	XSPECIALABORTBEHAVIOR : BOOL;
	LRABORTDEC : LREAL;
	LRABORTJERK : LREAL;
END_VAR
VAR_OUTPUT
	XERROR : BOOL;
	EERRORID : L_TB2P.L_IE1P_Error;
	XFUNBUSY : BOOL;
	XFUNDONE : BOOL;
	XFUNCOMMANDABORTED : BOOL;
	EFUNSTATEACT : L_TB2P.L_MC1P_ABC_State;
	ECONTROLMODE : L_TB2P.L_MC1P_ControlMode;
	XISHOMED : BOOL;
	XHWLIMITSWITCHNEG : BOOL;
	XHWLIMITSWITCHPOS : BOOL;
	XSWLIMITENABLED : BOOL;
	XSWLIMITSWITCHNEG : BOOL;
	XSWLIMITSWITCHPOS : BOOL;
	EAXISTYPE : L_TB2P.L_MC1P_DriveType;
	EAXISSTATE : L_TB2P.L_MC1P_AXIS_STATE;
	XSTOACTIVE : BOOL;
	XREADYFOROPERATION : BOOL;
	XOPERATIONENABLED : BOOL;
	XREADYFORMOTION : BOOL;
	XAXISWARNING : BOOL;
	XAXISERROR : BOOL;
	EAXISERRORID : L_TB2P.L_IE1P_Error;
	XDRIVEWARNING : BOOL;
	XDRIVEERROR : BOOL;
	DWDRIVEERRORID : DWORD;
	LRACTPOS : LREAL;
	LRACTVEL : LREAL;
	LRSETPOSOUT : LREAL;
	LRSETVELOUT : LREAL;
	LRACTFOLLOWINGERROR : LREAL;
	XINPOSITION : BOOL;
	XSTANDSTILLSETVELOCITY : BOOL;
	XSTANDSTILLACTVELOCITY : BOOL;
	XCONSTANTVELOCITY : BOOL;
	XACCELERATING : BOOL;
	XDECELERATING : BOOL;
	XDIRECTIONPOSITIVE : BOOL;
	XDIRECTIONNEGATIVE : BOOL;
	XAXISAVAILABLE : BOOL;
END_VAR
VAR_IN_OUT
	AXIS : AXIS_REF;
END_VAR
END_METHOD

METHOD GET_PAP : POINTER TO L_TB2P_scAP_TM_MotionControl
END_METHOD

METHOD GET_PDATA : POINTER TO L_TS2P_scData_TM_FlexCam
END_METHOD

METHOD GET_PDATASP : POINTER TO L_TS2P_scData_TM_FlexCam
END_METHOD

METHOD GET_PPAR : POINTER TO L_TB2P.L_TB2P_scPar_TM_MotionControl
END_METHOD

METHOD GET_PSF : POINTER TO L_TB2P_scSF_TM_MotionControl
END_METHOD

METHOD CAM
VAR_INPUT
	ITFTECHMODULE : L_TS2P_IFlexCam;
	XENABLE : BOOL;
	XSYNCCAM : BOOL;
	SCCAMTABLE : L_MC2P.MC_CAM_REF;
	LRCYCMASTERPOS : LREAL;
	LRCYCMASTERVEL : LREAL;
	LRCYCMASTERACC : LREAL;
	LRSLAVEPOS : LREAL;
	LRSLAVEVEL : LREAL;
	LRSLAVEACC : LREAL;
	EOFFSETMODEMASTER : L_TS2P_OffsetMode := L_TS2P_OffsetMode.x_zero;
	ESCALINGMODEMASTER : L_TS2P_ScalingMode := L_TS2P_ScalingMode.x_zero;
	EOFFSETMODESLAVE : L_TS2P_OffsetMode := L_TS2P_OffsetMode.x_zero;
	ESCALINGMODESLAVE : L_TS2P_ScalingMode := L_TS2P_ScalingMode.x_zero;
	LRSETOFFSETMASTER : LREAL;
	LRSETOFFSETSLAVE : LREAL;
	LRSETSCALINGMASTER : LREAL;
	LRSETSCALINGSLAVE : LREAL;
	LRPROFGENMASTERVEL : LREAL;
	LRPROFGENMASTERACC : LREAL;
	LRPROFGENMASTERDEC : LREAL;
	LRPROFGENMASTERJERK : LREAL;
	LRPROFGENSLAVEVEL : LREAL;
	LRPROFGENSLAVEACC : LREAL;
	LRPROFGENSLAVEDEC : LREAL;
	LRPROFGENSLAVEJERK : LREAL;
	XPERIODIC : BOOL;
	XCAMCHANGEINSTANT : BOOL;
	XMASTERABSOLUTE : BOOL;
	XSLAVEABSOLUTE : BOOL;
END_VAR
VAR_OUTPUT
	XERROR : BOOL;
	EERRORID : L_IE1P.L_IE1P_Error;
	LRSETPOSOUT : LREAL;
	LRSETVELOUT : LREAL;
	LRSETACCOUT : LREAL;
	LRSETXPOSOUT : LREAL;
	LRSETXVELOUT : LREAL;
	LRSETXACCOUT : LREAL;
	LRSETYPOSOUT : LREAL;
	LRSETYVELOUT : LREAL;
	LRSETYACCOUT : LREAL;
	XENDOFPROFILE : BOOL;
	LRSETOFFSETMASTEROUT : LREAL;
	LRSETOFFSETSLAVEOUT : LREAL;
	LRCONVERTMASTERTOXPOS : LREAL;
	LRCAMPROFILERPOSOUT : LREAL;
	LRCONVERTYTOSLAVEPOS : LREAL;
	XDONE : BOOL;
	XBUSY : BOOL;
END_VAR
END_METHOD

METHOD CAMSEQUENCER
VAR_INPUT
	ITFTECHMODULE : L_TS2P_IFlexCam;
	XENABLE : BOOL;
	XCAMSEQUENCER : BOOL;
	XENDOFPROFILEIN : BOOL;
	CAMTABLE1 : L_MC2P.MC_CAM_REF;
	CAMTABLE2 : L_MC2P.MC_CAM_REF;
	CAMTABLE3 : L_MC2P.MC_CAM_REF;
	CAMTABLE4 : L_MC2P.MC_CAM_REF;
	XCAMCHANGEINSTANT : BOOL;
	XLOADCAMTABLE : BOOL;
	WSETCAMTABLE : WORD;
	EMODE : L_TS2P_CamSequenceMode := L_TS2P_CamSequenceMode.CyclicCam1;
END_VAR
VAR_OUTPUT
	XERROR : BOOL;
	EERRORID : L_IE1P_Error;
	CAMTABLEOUT : L_MC2P.MC_CAM_REF;
	XCAMTABLEVALID : BOOL;
END_VAR
END_METHOD

METHOD CLUTCH
VAR_INPUT
	ITFTECHMODULE : L_TS2P_IFlexCam;
	XENABLE : BOOL;
	XCLUTCHCLOSE : BOOL;
	ECLUTCHINMODE : L_TS2P_ClutchInMode;
	ECLUTCHOUTMODE : L_TS2P_ClutchOutMode;
	EALLOWEDDIRECTION : L_TB2P_AllowedDirection;
	LRCLUTCHINDIST : LREAL;
	LRCLUTCHOUTDIST : LREAL;
	LRCLUTCHOUTPOSITION : LREAL;
	LRCYCLICMASTERPOS : LREAL;
	LRCYCLICMASTERVEL : LREAL;
	LRCYCLICMASTERACC : LREAL;
	LRCYCLICAXISPOS : LREAL;
	LRCYCLICAXISVEL : LREAL;
	LRCYCLICAXISACC : LREAL;
	ETRAVERSINGRANGE : L_MC1P_TraversingRange;
	LRCYCLELENGTH : LREAL;
END_VAR
VAR_OUTPUT
	XERROR : BOOL;
	EERRORID : L_IE1P.L_IE1P_Error;
	XBUSY : BOOL;
	XDONE : BOOL;
	XSYNCHRONISED : BOOL;
	XACCDECSYNC : BOOL;
	LRSETPOSOUT : LREAL;
	LRSETVELOUT : LREAL;
	LRSETACCOUT : LREAL;
END_VAR
END_METHOD

METHOD HALT : BOOL
VAR_INPUT
	ITFTECHMODULE : L_TS2P_IFlexCam;
	XEXECUTE : BOOL;
	LRDEC : LREAL := 100;
	LRJERK : LREAL := 0;
END_VAR
VAR_OUTPUT
	XBUSY : BOOL;
	XDONE : BOOL;
	XCOMMANDABORTED : BOOL;
END_VAR
VAR_IN_OUT
	AXIS : AXIS_REF;
END_VAR
END_METHOD

METHOD MOVETOPARKPOS : BOOL
VAR_INPUT
	ITFTECHMODULE : L_TS2P_IFlexCam;
	XEXECUTEMOVETOPARKPOS : BOOL;
	EMOVETOPARKPOSMODE : L_TS2P_CamStopMode;
	LRPARKPOSITION : LREAL := 180;
	EPOSITIONINGDIRECTION : L_TS2P_SyncDirection := L_TS2P_SyncDirection.PositiveDirection;
	LRPOSITIONINGVEL : LREAL := 10;
	LRPOSITIONINGACC : LREAL := 100;
	LRPOSITIONINGDEC : LREAL := 100;
	LRJERK : LREAL := 0;
END_VAR
VAR_OUTPUT
	XBUSY : BOOL;
	XDONE : BOOL;
	XCOMMANDABORTED : BOOL;
END_VAR
VAR_IN_OUT
	AXIS : AXIS_REF;
END_VAR
END_METHOD

METHOD POSITIONFOLLOWER
VAR_INPUT
	ITFTECHMODULE : L_TS2P_IFlexCam;
	XENABLE : BOOL;
	LRPOSITION : LREAL;
	LRVELOCITY : LREAL;
	LRACCELERATION : LREAL;
	ESETVALUEMODE : L_MC1P_SetValueMode;
END_VAR
VAR_OUTPUT
	XERROR : BOOL;
	EERRORID : L_IE1P.L_IE1P_Error;
	XBUSY : BOOL;
END_VAR
END_METHOD

METHOD SYNCIN
VAR_INPUT
	ITFTECHMODULE : L_TS2P_IFlexCam;
	XENABLE : BOOL;
	XSYNCIN : BOOL;
	XSYNCPOSRESTORE : BOOL;
	ESYNCMODE : L_TS2P_SyncInMode;
	ESYNCDIRECTION : L_TS2P_SyncDirection;
	LRSYNCVEL : LREAL;
	LRSYNCACC : LREAL;
	LRSYNCDEC : LREAL;
	LRSYNCJERK : LREAL;
	LRPARKPOSITION : LREAL;
	LRCYCLICMASTERPOS : LREAL;
	LRCYCLICMASTERVEL : LREAL;
	LRCYCLICMASTERACC : LREAL;
	LRCYCLICAXISPOS : LREAL;
	LRCYCLICAXISVEL : LREAL;
	LRCYCLICAXISACC : LREAL;
END_VAR
VAR_OUTPUT
	XERROR : BOOL;
	EERRORID : L_IE1P.L_IE1P_Error;
	XBUSY : BOOL;
	XDONE : BOOL;
	XSYNCHRONISED : BOOL;
	XACCDECSYNC : BOOL;
	LRSETPOSOUT : LREAL;
	LRSETVELOUT : LREAL;
	LRSETACCOUT : LREAL;
	LROFFSETSYNCPOS : LREAL;
END_VAR
VAR_IN_OUT
	AXIS : AXIS_REF;
END_VAR
END_METHOD

METHOD REQUESTINTERFACE : BOOL
VAR_INPUT
	ID : DINT;
	PITFUNKNOWN : POINTER TO L_UBUP.L_UBUP_IUnknown;
END_VAR
END_METHOD

METHOD CALLFUNCTION
VAR_INPUT
	UIINPUTDATAIDX : UINT;
	UIOUTPUTDATAIDX : UINT;
END_VAR
END_METHOD

METHOD COPYINPUTS : BOOL
VAR_INPUT
	IDX : WORD;
END_VAR
END_METHOD

METHOD COPYOUTPUTS : BOOL
VAR_INPUT
	IDX : WORD;
END_VAR
END_METHOD

METHOD FUNCTIONWASCALLEDTWICE : BOOL
VAR_INPUT
	IDX : WORD;
END_VAR
END_METHOD

METHOD HANDLESTANDARDCALL : BOOL
END_METHOD

METHOD SYNCOUTPUTS
VAR_INPUT
	UICOPYOUTPUTFROMIDX : UINT;
	UICOPYOUTPUTTOIDX : UINT;
END_VAR
END_METHOD

METHOD FB_INIT : BOOL
VAR_INPUT
	BINITRETAINS : BOOL;
	BINCOPYCODE : BOOL;
END_VAR
END_METHOD

METHOD CALL_INTERNALCTRL
END_METHOD

METHOD GET_INTERNCAMTABLE : MC_CAM_REF
END_METHOD

METHOD GET_LRCAMXEND : LREAL
END_METHOD

METHOD GET_LRCAMXSTART : LREAL
END_METHOD

METHOD GET_LRCAMYEND : LREAL
END_METHOD

METHOD GET_LRCAMYSTART : LREAL
END_METHOD

METHOD GET_STCAMNAME : STRING
END_METHOD

METHOD GET_XCOMMUNICATION : BOOL
END_METHOD

(* ---- L_TS2P_FLEXCAMSTATE.fb ---- *)
FUNCTION_BLOCK L_TS2P_FLEXCAMSTATE EXTENDS L_TB2P_TechModuleBase
VAR_INPUT
	XENABLE : BOOL;
	XENABLEOPERATION : BOOL;
	XRESETERROR : BOOL;
	XQSPAPPLICATION : BOOL;
	XABORT : BOOL;
	XJOGPOS : BOOL;
	XJOGNEG : BOOL;
	XHOMEEXECUTE : BOOL;
	LROVERRIDE : LREAL := 1;
	SCCTRLBASICMOTION : L_TB2P_scCtrlBasicMotion;
	SCPAR : L_TS2P_scPar_FlexCamState;
	SCACCESSPOINTS : L_TS2P_scAP_FlexCamState;
	MASTERVALUES : L_MC1P_IAXIS_REF_MASTERVALUES;
	XSYNCIN : BOOL;
	XCAMCHANGEINSTANT : BOOL;
	LRSETOFFSETPOSX : LREAL;
	LRSETOFFSETPOSY : LREAL;
	LRSETSCALINGX : LREAL := 1;
	LRSETSCALINGY : LREAL := 1;
	CAMTABLE1 : MC_CAM_REF;
	CAMTABLE2 : MC_CAM_REF;
	CAMTABLE3 : MC_CAM_REF;
	CAMTABLE4 : MC_CAM_REF;
	WSETCAMTABLE : WORD := 1;
	XCAMSEQUENCER : BOOL;
END_VAR
VAR_OUTPUT
	XREADYFOROPERATION : BOOL;
	XOPERATIONENABLED : BOOL;
	XREADYFORMOTION : BOOL;
	XERROR : BOOL;
	XWARNING : BOOL;
	EERRORID : L_IE1P_Error;
	XSTOACTIVE : BOOL;
	XQSPACTIVE : BOOL;
	XABORTBUSY : BOOL;
	XABORTDONE : BOOL;
	XJOGGINGBUSY : BOOL;
	XHOMINGBUSY : BOOL;
	XHOMINGDONE : BOOL;
	XISHOMED : BOOL;
	ETMSTATE : L_TB2P_States := L_TB2P_States.DISABLED;
	SCSTATUSBASICMOTION : L_TB2P_scStatusBasicMotion;
	LRACTVEL : LREAL;
	LRSETVELOUT : LREAL;
	LRACTPOS : LREAL;
	LRSETPOSOUT : LREAL;
	LRACTFOLLOWINGERROR : LREAL;
	SCSIGNALFLOW : L_TS2P_scSF_FlexCamState;
	XSYNCHRONISED : BOOL;
	XACCDECSYNC : BOOL;
	XCAMMINGBUSY : BOOL;
	XENDOFPROFILE : BOOL;
	LROFFSETPOSX : LREAL;
	LROFFSETPOSY : LREAL;
	WACTIVECAMTABLE : WORD;
	XCAMSEQUENCERACTIVE : BOOL;
END_VAR
VAR_IN_OUT
	AXIS : AXIS_REF;
END_VAR
VAR
	TM_INT : L_TS2P_TM_FlexCamState := STRUCT(ModuleHandler := ModuleHandler);
	SCPAR_INT : L_TS2P_scPar_FlexCamState;
	_UICALLMFUNIDXINPUT : UINT := 1;
	_UICALLMFUNIDXOUTPUT : UINT := 1;
	_MCCALL : L_UM1P_MCCall;
	_ASCINPUT : ARRAY [1.._MCCall.c_BufferDepthInput] OF L_TS2P_FlexCamStateIn;
	_ASCOUTPUT : ARRAY [1.._MCCall.c_BufferDepthOutput] OF L_TS2P_FlexCamStateOut;
	_ASCPARCORE : ARRAY [1.._MCCall.c_BufferDepthInput] OF L_TS2P_scPar_FlexCamState;
	_ASCACCESSPOINTSCORE : ARRAY [1.._MCCall.c_BufferDepthInput] OF L_TS2P_scAp_FlexCamState;
	_ASCSIGNALFLOWCORE : ARRAY [1.._MCCall.c_BufferDepthOutput] OF L_TS2P_scSF_FlexCamState;
	_SCINPUTVISU : L_TS2P_FlexCamStateIn;
	_PSCINPUTVISU : POINTER TO L_TS2P_FlexCamStateIn := ADR(_scInputVisu);
	_PSCOUTPUTVISU : POINTER TO L_TS2P_FlexCamStateOut := ADR(_ascOutput[1]);
	_PSCPARVISU : POINTER TO L_TS2P_scPar_FlexCamState := ADR(scPar_int);
	ITFITECHMODULEINTERNAL : L_TB2P_ITechModuleInternal;
	LRJERKDEC : LREAL;
	LRJOGGINGJERKDEC : LREAL;
	REMAININGTIMEOFPROFILE : LREAL;
	REMAININGTIMEOFPROFILEAVAILABLE : BOOL;
END_VAR
END_FUNCTION_BLOCK

METHOD GET_INTERNCAMTABLE : MC_CAM_REF
END_METHOD

METHOD GET_LRCAMXEND : LREAL
END_METHOD

METHOD GET_LRCAMXSTART : LREAL
END_METHOD

METHOD GET_LRCAMYEND : LREAL
END_METHOD

METHOD GET_LRCAMYSTART : LREAL
END_METHOD

METHOD GET_STCAMNAME : STRING
END_METHOD

METHOD GET_XCOMMUNICATION : BOOL
END_METHOD

METHOD GET_PAP : POINTER TO L_TB2P_scAP_TM_MotionControl
END_METHOD

METHOD GET_PPAR : POINTER TO L_TB2P_scPar_TM_MotionControl
END_METHOD

METHOD GET_PSF : POINTER TO L_TB2P_scSF_TM_MotionControl
END_METHOD

METHOD CALLFUNCTION
VAR_INPUT
	UIINPUTDATAIDX : UINT;
	UIOUTPUTDATAIDX : UINT;
END_VAR
END_METHOD

METHOD COPYINPUTS : BOOL
VAR_INPUT
	IDX : WORD;
END_VAR
END_METHOD

METHOD COPYOUTPUTS : BOOL
VAR_INPUT
	IDX : WORD;
END_VAR
END_METHOD

METHOD FUNCTIONWASCALLEDTWICE : BOOL
VAR_INPUT
	IDX : WORD;
END_VAR
END_METHOD

METHOD HANDLESTANDARDCALL : BOOL
END_METHOD

METHOD SYNCOUTPUTS
VAR_INPUT
	UICOPYOUTPUTFROMIDX : UINT;
	UICOPYOUTPUTTOIDX : UINT;
END_VAR
END_METHOD

METHOD CALL_INTERNALCTRL
END_METHOD
